(* IEC 61131-3 sources: BODAS-HelloWorld/st/bodas_rc18_12_40/plc_logic/application/02_easyconfig/dsm_easyconfig/structure (part 2) *)

(* ---- dfc_bds_tiinrow0x8b02-DFC_bds_TiInRow0x8B02.st ---- *)
(* --- Interface --- *)
{attribute 'external_name' := 'cmp_rts_DFC_bds_TiInRow0x8B02'}
TYPE DFC_bds_TiInRow0x8B02 : STRUCT
		DTC            : UDINT := 16#8B0200;
		DFCid          : UINT  := 102;
		debounceMethod : USINT := TIME_IN_ROW;
	END_STRUCT
END_TYPE

(* ---- dfc_bds_tiinrow0x8b03-DFC_bds_TiInRow0x8B03.st ---- *)
(* --- Interface --- *)
{attribute 'external_name' := 'cmp_rts_DFC_bds_TiInRow0x8B03'}
TYPE DFC_bds_TiInRow0x8B03 : STRUCT
		DTC            : UDINT := 16#8B0300;
		DFCid          : UINT  := 103;
		debounceMethod : USINT := TIME_IN_ROW;
	END_STRUCT
END_TYPE

(* ---- dfc_bds_tiupdwn0x8a01-DFC_bds_TiUpDwn0x8A01.st ---- *)
(* --- Interface --- *)
{attribute 'external_name' := 'cmp_rts_DFC_bds_TiUpDwn0x8A01'}
TYPE DFC_bds_TiUpDwn0x8A01 : STRUCT
		DTC            : UDINT := 16#8A0100;
		DFCid          : UINT  := 206;
		debounceMethod : USINT := TIME_UP_DOWN;
	END_STRUCT
END_TYPE

(* ---- dfc_bds_tiupdwn0x8a02-DFC_bds_TiUpDwn0x8A02.st ---- *)
(* --- Interface --- *)
{attribute 'external_name' := 'cmp_rts_DFC_bds_TiUpDwn0x8A02'}
TYPE DFC_bds_TiUpDwn0x8A02 : STRUCT
		DTC            : UDINT := 16#8A0200;
		DFCid          : UINT  := 207;
		debounceMethod : USINT := TIME_UP_DOWN;
	END_STRUCT
END_TYPE

(* ---- dfc_bds_tiupdwn0x8a03-DFC_bds_TiUpDwn0x8A03.st ---- *)
(* --- Interface --- *)
{attribute 'external_name' := 'cmp_rts_DFC_bds_TiUpDwn0x8A03'}
TYPE DFC_bds_TiUpDwn0x8A03 : STRUCT
		DTC            : UDINT := 16#8A0300;
		DFCid          : UINT  := 208;
		debounceMethod : USINT := TIME_UP_DOWN;
	END_STRUCT
END_TYPE

(* ---- dfc_can_e_timeout-DFC_CAN_E_TIMEOUT.st ---- *)
(* --- Interface --- *)
{attribute 'external_name' := 'cmp_rts_DFC_CAN_E_TIMEOUT'}
TYPE DFC_CAN_E_TIMEOUT : STRUCT
		DTC            : UDINT := 16#094200;
		DFCid          : UINT  := 1165;
		debounceMethod : USINT := NO_DEBOUNCE;
	END_STRUCT
END_TYPE

(* ---- dfc_cansm_e_bus_off_network_0-DFC_CANSM_E_BUS_OFF_NETWORK_0.st ---- *)
(* --- Interface --- *)
{attribute 'external_name' := 'cmp_rts_DFC_CANSM_E_BUS_OFF_NETWORK_0'}
TYPE DFC_CANSM_E_BUS_OFF_NETWORK_0 : STRUCT
		DTC            : UDINT := 16#104C00;
		DFCid          : UINT  := 1160;
		debounceMethod : USINT := NO_DEBOUNCE;
	END_STRUCT
END_TYPE

(* ---- dfc_cansm_e_bus_off_network_1-DFC_CANSM_E_BUS_OFF_NETWORK_1.st ---- *)
(* --- Interface --- *)
{attribute 'external_name' := 'cmp_rts_DFC_CANSM_E_BUS_OFF_NETWORK_1'}
TYPE DFC_CANSM_E_BUS_OFF_NETWORK_1 : STRUCT
		DTC            : UDINT := 16#104D00;
		DFCid          : UINT  := 1161;
		debounceMethod : USINT := NO_DEBOUNCE;
	END_STRUCT
END_TYPE

(* ---- dfc_cansm_e_bus_off_network_2-DFC_CANSM_E_BUS_OFF_NETWORK_2.st ---- *)
(* --- Interface --- *)
{attribute 'external_name' := 'cmp_rts_DFC_CANSM_E_BUS_OFF_NETWORK_2'}
TYPE DFC_CANSM_E_BUS_OFF_NETWORK_2 : STRUCT
		DTC            : UDINT := 16#104E00;
		DFCid          : UINT  := 1162;
		debounceMethod : USINT := NO_DEBOUNCE;
	END_STRUCT
END_TYPE

(* ---- dfc_cansm_e_bus_off_network_3-DFC_CANSM_E_BUS_OFF_NETWORK_3.st ---- *)
(* --- Interface --- *)
{attribute 'external_name' := 'cmp_rts_DFC_CANSM_E_BUS_OFF_NETWORK_3'}
TYPE DFC_CANSM_E_BUS_OFF_NETWORK_3 : STRUCT
		DTC            : UDINT := 16#104F00;
		DFCid          : UINT  := 1163;
		debounceMethod : USINT := NO_DEBOUNCE;
	END_STRUCT
END_TYPE

(* ---- dfc_cantrcv_e_no_trcv_control_0-DFC_CANTRCV_E_NO_TRCV_CONTROL_0.st ---- *)
(* --- Interface --- *)
{attribute 'external_name' := 'cmp_rts_DFC_CANTRCV_E_NO_TRCV_CONTROL_0'}
TYPE DFC_CANTRCV_E_NO_TRCV_CONTROL_0 : STRUCT
		DTC            : UDINT := 16#094000;
		DFCid          : UINT  := 1164;
		debounceMethod : USINT := NO_DEBOUNCE;
	END_STRUCT
END_TYPE

(* ---- dfc_com_numwhlincfrtleft-DFC_Com_numWhlIncFrtLeft.st ---- *)
(* --- Interface --- *)
{attribute 'external_name' := 'cmp_rts_DFC_Com_numWhlIncFrtLeft'}
TYPE DFC_Com_numWhlIncFrtLeft : STRUCT
		DTC : UDINT := 16#103A00;
	END_STRUCT
END_TYPE

(* ---- dfc_com_stwhlsensrrrht-DFC_Com_stWhlSensRrRht.st ---- *)
(* --- Interface --- *)
{attribute 'external_name' := 'cmp_rts_DFC_Com_stWhlSensRrRht'}
TYPE DFC_Com_stWhlSensRrRht : STRUCT
		DTC : UDINT := 16#103B00;
	END_STRUCT
END_TYPE

(* ---- dfc_com_trqclthtcsdcsdes-DFC_Com_trqClthTCSDCSDes.st ---- *)
(* --- Interface --- *)
{attribute 'external_name' := 'cmp_rts_DFC_Com_trqClthTCSDCSDes'}
TYPE DFC_Com_trqClthTCSDCSDes : STRUCT
		DTC : UDINT := 16#103C00;
	END_STRUCT
END_TYPE

(* ---- dfc_com_vwhlrrl-DFC_Com_vWhlRrL.st ---- *)
(* --- Interface --- *)
{attribute 'external_name' := 'cmp_rts_DFC_Com_vWhlRrL'}
TYPE DFC_Com_vWhlRrL : STRUCT
		DTC : UDINT := 16#103D00;
	END_STRUCT
END_TYPE

(* ---- dfc_comchksacc_06-DFC_ComChksACC_06.st ---- *)
(* --- Interface --- *)
{attribute 'external_name' := 'cmp_rts_DFC_ComChksACC_06'}
TYPE DFC_ComChksACC_06 : STRUCT
		DTC : UDINT := 16#101600;
	END_STRUCT
END_TYPE

(* ---- dfc_comchksbms_01-DFC_ComChksBMS_01.st ---- *)
(* --- Interface --- *)
{attribute 'external_name' := 'cmp_rts_DFC_ComChksBMS_01'}
TYPE DFC_ComChksBMS_01 : STRUCT
		DTC : UDINT := 16#101700;
	END_STRUCT
END_TYPE

(* ---- dfc_comchksesp_02-DFC_ComChksESP_02.st ---- *)
(* --- Interface --- *)
{attribute 'external_name' := 'cmp_rts_DFC_ComChksESP_02'}
TYPE DFC_ComChksESP_02 : STRUCT
		DTC : UDINT := 16#101800;
	END_STRUCT
END_TYPE

(* ---- dfc_comchksesp_05-DFC_ComChksESP_05.st ---- *)
(* --- Interface --- *)
{attribute 'external_name' := 'cmp_rts_DFC_ComChksESP_05'}
TYPE DFC_ComChksESP_05 : STRUCT
		DTC : UDINT := 16#101900;
	END_STRUCT
END_TYPE

(* ---- dfc_comchksesp_07-DFC_ComChksESP_07.st ---- *)
(* --- Interface --- *)
{attribute 'external_name' := 'cmp_rts_DFC_ComChksESP_07'}
TYPE DFC_ComChksESP_07 : STRUCT
		DTC : UDINT := 16#101A00;
	END_STRUCT
END_TYPE

(* ---- dfc_comchksesp_10-DFC_ComChksESP_10.st ---- *)
(* --- Interface --- *)
{attribute 'external_name' := 'cmp_rts_DFC_ComChksESP_10'}
TYPE DFC_ComChksESP_10 : STRUCT
		DTC : UDINT := 16#101B00;
	END_STRUCT
END_TYPE

(* ---- dfc_comchksesp_19-DFC_ComChksESP_19.st ---- *)
(* --- Interface --- *)
{attribute 'external_name' := 'cmp_rts_DFC_ComChksESP_19'}
TYPE DFC_ComChksESP_19 : STRUCT
		DTC : UDINT := 16#101C00;
	END_STRUCT
END_TYPE

(* ---- dfc_comchksesp_20-DFC_ComChksESP_20.st ---- *)
(* --- Interface --- *)
{attribute 'external_name' := 'cmp_rts_DFC_ComChksESP_20'}
TYPE DFC_ComChksESP_20 : STRUCT
		DTC : UDINT := 16#101D00;
	END_STRUCT
END_TYPE

(* ---- dfc_comchksesp_21-DFC_ComChksESP_21.st ---- *)
(* --- Interface --- *)
{attribute 'external_name' := 'cmp_rts_DFC_ComChksESP_21'}
TYPE DFC_ComChksESP_21 : STRUCT
		DTC : UDINT := 16#101E00;
	END_STRUCT
END_TYPE

(* ---- dfc_comchksklemmen_status_01-DFC_ComChksKlemmen_Status_01.st ---- *)
(* --- Interface --- *)
{attribute 'external_name' := 'cmp_rts_DFC_ComChksKlemmen_Status_01'}
TYPE DFC_ComChksKlemmen_Status_01 : STRUCT
		DTC : UDINT := 16#103800;
	END_STRUCT
END_TYPE

(* ---- dfc_comcntacc_06-DFC_ComCntACC_06.st ---- *)
(* --- Interface --- *)
{attribute 'external_name' := 'cmp_rts_DFC_ComCntACC_06'}
TYPE DFC_ComCntACC_06 : STRUCT
		DTC : UDINT := 16#101F00;
	END_STRUCT
END_TYPE

(* ---- dfc_comcntbms_01-DFC_ComCntBMS_01.st ---- *)
(* --- Interface --- *)
{attribute 'external_name' := 'cmp_rts_DFC_ComCntBMS_01'}
TYPE DFC_ComCntBMS_01 : STRUCT
		DTC : UDINT := 16#102000;
	END_STRUCT
END_TYPE

(* ---- dfc_comcntesp_02-DFC_ComCntESP_02.st ---- *)
(* --- Interface --- *)
{attribute 'external_name' := 'cmp_rts_DFC_ComCntESP_02'}
TYPE DFC_ComCntESP_02 : STRUCT
		DTC : UDINT := 16#102100;
	END_STRUCT
END_TYPE

(* ---- dfc_comcntesp_05-DFC_ComCntESP_05.st ---- *)
(* --- Interface --- *)
{attribute 'external_name' := 'cmp_rts_DFC_ComCntESP_05'}
TYPE DFC_ComCntESP_05 : STRUCT
		DTC : UDINT := 16#102200;
	END_STRUCT
END_TYPE

(* ---- dfc_comcntesp_07-DFC_ComCntESP_07.st ---- *)
(* --- Interface --- *)
{attribute 'external_name' := 'cmp_rts_DFC_ComCntESP_07'}
TYPE DFC_ComCntESP_07 : STRUCT
		DTC : UDINT := 16#102300;
	END_STRUCT
END_TYPE

(* ---- dfc_comcntesp_10-DFC_ComCntESP_10.st ---- *)
(* --- Interface --- *)
{attribute 'external_name' := 'cmp_rts_DFC_ComCntESP_10'}
TYPE DFC_ComCntESP_10 : STRUCT
		DTC : UDINT := 16#102400;
	END_STRUCT
END_TYPE

(* ---- dfc_comcntesp_19-DFC_ComCntESP_19.st ---- *)
(* --- Interface --- *)
{attribute 'external_name' := 'cmp_rts_DFC_ComCntESP_19'}
TYPE DFC_ComCntESP_19 : STRUCT
		DTC : UDINT := 16#102500;
	END_STRUCT
END_TYPE

(* ---- dfc_comcntesp_20-DFC_ComCntESP_20.st ---- *)
(* --- Interface --- *)
{attribute 'external_name' := 'cmp_rts_DFC_ComCntESP_20'}
TYPE DFC_ComCntESP_20 : STRUCT
		DTC : UDINT := 16#102600;
	END_STRUCT
END_TYPE

(* ---- dfc_comcntesp_21-DFC_ComCntESP_21.st ---- *)
(* --- Interface --- *)
{attribute 'external_name' := 'cmp_rts_DFC_ComCntESP_21'}
TYPE DFC_ComCntESP_21 : STRUCT
		DTC : UDINT := 16#102700;
	END_STRUCT
END_TYPE

(* ---- dfc_comcntklemmen_status_01-DFC_ComCntKlemmen_Status_01.st ---- *)
(* --- Interface --- *)
{attribute 'external_name' := 'cmp_rts_DFC_ComCntKlemmen_Status_01'}
TYPE DFC_ComCntKlemmen_Status_01 : STRUCT
		DTC : UDINT := 16#103900;
	END_STRUCT
END_TYPE

(* ---- dfc_comdlcacc_06-DFC_ComDlcACC_06.st ---- *)
(* --- Interface --- *)
{attribute 'external_name' := 'cmp_rts_DFC_ComDlcACC_06'}
TYPE DFC_ComDlcACC_06 : STRUCT
		DTC : UDINT := 16#102800;
	END_STRUCT
END_TYPE

(* ---- dfc_comdlcesp_02-DFC_ComDlcESP_02.st ---- *)
(* --- Interface --- *)
{attribute 'external_name' := 'cmp_rts_DFC_ComDlcESP_02'}
TYPE DFC_ComDlcESP_02 : STRUCT
		DTC : UDINT := 16#102900;
	END_STRUCT
END_TYPE

(* ---- dfc_comdlcesp_05-DFC_ComDlcESP_05.st ---- *)
(* --- Interface --- *)
{attribute 'external_name' := 'cmp_rts_DFC_ComDlcESP_05'}
TYPE DFC_ComDlcESP_05 : STRUCT
		DTC : UDINT := 16#102A00;
	END_STRUCT
END_TYPE

(* ---- dfc_comdlcesp_07-DFC_ComDlcESP_07.st ---- *)
(* --- Interface --- *)
{attribute 'external_name' := 'cmp_rts_DFC_ComDlcESP_07'}
TYPE DFC_ComDlcESP_07 : STRUCT
		DTC : UDINT := 16#102B00;
	END_STRUCT
END_TYPE

(* ---- dfc_comdlcesp_10-DFC_ComDlcESP_10.st ---- *)
(* --- Interface --- *)
{attribute 'external_name' := 'cmp_rts_DFC_ComDlcESP_10'}
TYPE DFC_ComDlcESP_10 : STRUCT
		DTC : UDINT := 16#102C00;
	END_STRUCT
END_TYPE

(* ---- dfc_comdlcesp_19-DFC_ComDlcESP_19.st ---- *)
(* --- Interface --- *)
{attribute 'external_name' := 'cmp_rts_DFC_ComDlcESP_19'}
TYPE DFC_ComDlcESP_19 : STRUCT
		DTC : UDINT := 16#102D00;
	END_STRUCT
END_TYPE

(* ---- dfc_comdlcesp_20-DFC_ComDlcESP_20.st ---- *)
(* --- Interface --- *)
{attribute 'external_name' := 'cmp_rts_DFC_ComDlcESP_20'}
TYPE DFC_ComDlcESP_20 : STRUCT
		DTC : UDINT := 16#102E00;
	END_STRUCT
END_TYPE

(* ---- dfc_comdlcesp_21-DFC_ComDlcESP_21.st ---- *)
(* --- Interface --- *)
{attribute 'external_name' := 'cmp_rts_DFC_ComDlcESP_21'}
TYPE DFC_ComDlcESP_21 : STRUCT
		DTC : UDINT := 16#102F00;
	END_STRUCT
END_TYPE

(* ---- dfc_comm_e_net_start_ind_channel_0-DFC_COMM_E_NET_START_IND_CHANNEL_0.st ---- *)
(* --- Interface --- *)
{attribute 'external_name' := 'cmp_rts_DFC_COMM_E_NET_START_IND_CHANNEL_0'}
TYPE DFC_COMM_E_NET_START_IND_CHANNEL_0 : STRUCT
		DTC            : UDINT := 16#105000;
		DFCid          : UINT  := 1166;
		debounceMethod : USINT := NO_DEBOUNCE;
	END_STRUCT
END_TYPE

(* ---- dfc_comm_e_net_start_ind_channel_1-DFC_COMM_E_NET_START_IND_CHANNEL_1.st ---- *)
(* --- Interface --- *)
{attribute 'external_name' := 'cmp_rts_DFC_COMM_E_NET_START_IND_CHANNEL_1'}
TYPE DFC_COMM_E_NET_START_IND_CHANNEL_1 : STRUCT
		DTC            : UDINT := 16#105100;
		DFCid          : UINT  := 1167;
		debounceMethod : USINT := NO_DEBOUNCE;
	END_STRUCT
END_TYPE

(* ---- dfc_comm_e_net_start_ind_channel_2-DFC_COMM_E_NET_START_IND_CHANNEL_2.st ---- *)
(* --- Interface --- *)
{attribute 'external_name' := 'cmp_rts_DFC_COMM_E_NET_START_IND_CHANNEL_2'}
TYPE DFC_COMM_E_NET_START_IND_CHANNEL_2 : STRUCT
		DTC            : UDINT := 16#105200;
		DFCid          : UINT  := 1168;
		debounceMethod : USINT := NO_DEBOUNCE;
	END_STRUCT
END_TYPE

(* ---- dfc_comm_e_net_start_ind_channel_3-DFC_COMM_E_NET_START_IND_CHANNEL_3.st ---- *)
(* --- Interface --- *)
{attribute 'external_name' := 'cmp_rts_DFC_COMM_E_NET_START_IND_CHANNEL_3'}
TYPE DFC_COMM_E_NET_START_IND_CHANNEL_3 : STRUCT
		DTC            : UDINT := 16#105300;
		DFCid          : UINT  := 1169;
		debounceMethod : USINT := NO_DEBOUNCE;
	END_STRUCT
END_TYPE

(* ---- dfc_comm_e_net_start_ind_channel_4-DFC_COMM_E_NET_START_IND_CHANNEL_4.st ---- *)
(* --- Interface --- *)
{attribute 'external_name' := 'cmp_rts_DFC_COMM_E_NET_START_IND_CHANNEL_4'}
TYPE DFC_COMM_E_NET_START_IND_CHANNEL_4 : STRUCT
		DTC            : UDINT := 16#105400;
		DFCid          : UINT  := 1170;
		debounceMethod : USINT := NO_DEBOUNCE;
	END_STRUCT
END_TYPE

(* ---- dfc_comm_e_net_start_ind_channel_5-DFC_COMM_E_NET_START_IND_CHANNEL_5.st ---- *)
(* --- Interface --- *)
{attribute 'external_name' := 'cmp_rts_DFC_COMM_E_NET_START_IND_CHANNEL_5'}
TYPE DFC_COMM_E_NET_START_IND_CHANNEL_5 : STRUCT
		DTC            : UDINT := 16#105500;
		DFCid          : UINT  := 1171;
		debounceMethod : USINT := NO_DEBOUNCE;
	END_STRUCT
END_TYPE

(* ---- dfc_comtoutacc_06-DFC_ComTOutACC_06.st ---- *)
(* --- Interface --- *)
{attribute 'external_name' := 'cmp_rts_DFC_ComTOutACC_06'}
TYPE DFC_ComTOutACC_06 : STRUCT
		DTC : UDINT := 16#103000;
	END_STRUCT
END_TYPE

(* ---- dfc_comtoutesp_02-DFC_ComTOutESP_02.st ---- *)
(* --- Interface --- *)
{attribute 'external_name' := 'cmp_rts_DFC_ComTOutESP_02'}
TYPE DFC_ComTOutESP_02 : STRUCT
		DTC : UDINT := 16#103100;
	END_STRUCT
END_TYPE

(* ---- dfc_comtoutesp_05-DFC_ComTOutESP_05.st ---- *)
(* --- Interface --- *)
{attribute 'external_name' := 'cmp_rts_DFC_ComTOutESP_05'}
TYPE DFC_ComTOutESP_05 : STRUCT
		DTC : UDINT := 16#103200;
	END_STRUCT
END_TYPE

(* ---- dfc_comtoutesp_07-DFC_ComTOutESP_07.st ---- *)
(* --- Interface --- *)
{attribute 'external_name' := 'cmp_rts_DFC_ComTOutESP_07'}
TYPE DFC_ComTOutESP_07 : STRUCT
		DTC : UDINT := 16#103300;
	END_STRUCT
END_TYPE

(* ---- dfc_comtoutesp_10-DFC_ComTOutESP_10.st ---- *)
(* --- Interface --- *)
{attribute 'external_name' := 'cmp_rts_DFC_ComTOutESP_10'}
TYPE DFC_ComTOutESP_10 : STRUCT
		DTC : UDINT := 16#103400;
	END_STRUCT
END_TYPE

(* ---- dfc_comtoutesp_19-DFC_ComTOutESP_19.st ---- *)
(* --- Interface --- *)
{attribute 'external_name' := 'cmp_rts_DFC_ComTOutESP_19'}
TYPE DFC_ComTOutESP_19 : STRUCT
		DTC : UDINT := 16#103500;
	END_STRUCT
END_TYPE

(* ---- dfc_comtoutesp_20-DFC_ComTOutESP_20.st ---- *)
(* --- Interface --- *)
{attribute 'external_name' := 'cmp_rts_DFC_ComTOutESP_20'}
TYPE DFC_ComTOutESP_20 : STRUCT
		DTC : UDINT := 16#103600;
	END_STRUCT
END_TYPE

(* ---- dfc_comtoutesp_21-DFC_ComTOutESP_21.st ---- *)
(* --- Interface --- *)
{attribute 'external_name' := 'cmp_rts_DFC_ComTOutESP_21'}
TYPE DFC_ComTOutESP_21 : STRUCT
		DTC : UDINT := 16#103700;
	END_STRUCT
END_TYPE

(* ---- dfc_devlibbattuhi-DFC_DevLibBattUHi.st ---- *)
(* --- Interface --- *)
{attribute 'external_name' := 'cmp_rts_DFC_DevLibBattUHi'}
TYPE DFC_DevLibBattUHi : STRUCT
		DTC            : UDINT := 16#092300;
		DFCid          : UINT  := 104;
		debounceMethod : USINT := TIME_UP_DOWN;
	END_STRUCT
END_TYPE

(* ---- dfc_devlibbattulo-DFC_DevLibBattULo.st ---- *)
(* --- Interface --- *)
{attribute 'external_name' := 'cmp_rts_DFC_DevLibBattULo'}
TYPE DFC_DevLibBattULo : STRUCT
		DTC            : UDINT := 16#092400;
		DFCid          : UINT  := 105;
		debounceMethod : USINT := TIME_UP_DOWN;
	END_STRUCT
END_TYPE

(* ---- dfc_dsmdummy-DFC_DSMDummy.st ---- *)
(* --- Interface --- *)
{attribute 'external_name' := 'cmp_rts_DFC_DSMDummy'}
TYPE DFC_DSMDummy : STRUCT
		DTC            : UDINT := 16#100F00;
		DFCid          : UINT  := 720;
		debounceMethod : USINT := NO_DEBOUNCE;
	END_STRUCT
END_TYPE

(* ---- dfc_lin_e_timeout-DFC_LIN_E_TIMEOUT.st ---- *)
(* --- Interface --- *)
{attribute 'external_name' := 'cmp_rts_DFC_LIN_E_TIMEOUT'}
TYPE DFC_LIN_E_TIMEOUT : STRUCT
		DTC            : UDINT := 16#094100;
		DFCid          : UINT  := 1172;
		debounceMethod : USINT := NO_DEBOUNCE;
	END_STRUCT
END_TYPE

(* ---- dfc_mocsopico-DFC_MoCSOPICO.st ---- *)
(* --- Interface --- *)
{attribute 'external_name' := 'cmp_rts_DFC_MoCSOPICO'}
TYPE DFC_MoCSOPICO : STRUCT
		DTC            : UDINT := 16#106000;
		DFCid          : UINT  := 1296;
		debounceMethod : USINT := NATIVE;
	END_STRUCT
END_TYPE

(* ---- dfc_mofvarpostbldsel-DFC_MoFVarPostBldSel.st ---- *)
(* --- Interface --- *)
{attribute 'external_name' := 'cmp_rts_DFC_MoFVarPostBldSel'}
TYPE DFC_MoFVarPostBldSel : STRUCT
		DTC            : UDINT := 16#098900;
		DFCid          : UINT  := 1297;
		debounceMethod : USINT := NATIVE;
	END_STRUCT
END_TYPE

(* ---- dfc_mosysctrlreini-DFC_MoSysCtrlReIni.st ---- *)
(* --- Interface --- *)
{attribute 'external_name' := 'cmp_rts_DFC_MoSysCtrlReIni'}
TYPE DFC_MoSysCtrlReIni : STRUCT
		DTC            : UDINT := 16#106100;
		DFCid          : UINT  := 1298;
		debounceMethod : USINT := NATIVE;
	END_STRUCT
END_TYPE

(* ---- dfc_moxemm_smu_alm0_0-DFC_MOXEMM_SMU_ALM0_0.st ---- *)
(* --- Interface --- *)
{attribute 'external_name' := 'cmp_rts_DFC_MOXEMM_SMU_ALM0_0'}
TYPE DFC_MOXEMM_SMU_ALM0_0 : STRUCT
		DTC            : UDINT := 16#106200;
		DFCid          : UINT  := 1185;
		debounceMethod : USINT := NATIVE;
	END_STRUCT
END_TYPE

(* ---- dfc_moxemm_smu_alm0_1-DFC_MOXEMM_SMU_ALM0_1.st ---- *)
(* --- Interface --- *)
{attribute 'external_name' := 'cmp_rts_DFC_MOXEMM_SMU_ALM0_1'}
TYPE DFC_MOXEMM_SMU_ALM0_1 : STRUCT
		DTC            : UDINT := 16#106300;
		DFCid          : UINT  := 1186;
		debounceMethod : USINT := NATIVE;
	END_STRUCT
END_TYPE

(* ---- dfc_moxemm_smu_alm0_10-DFC_MOXEMM_SMU_ALM0_10.st ---- *)
(* --- Interface --- *)
{attribute 'external_name' := 'cmp_rts_DFC_MOXEMM_SMU_ALM0_10'}
TYPE DFC_MOXEMM_SMU_ALM0_10 : STRUCT
		DTC            : UDINT := 16#106900;
		DFCid          : UINT  := 1187;
		debounceMethod : USINT := NATIVE;
	END_STRUCT
END_TYPE

(* ---- dfc_moxemm_smu_alm0_11-DFC_MOXEMM_SMU_ALM0_11.st ---- *)
(* --- Interface --- *)
{attribute 'external_name' := 'cmp_rts_DFC_MOXEMM_SMU_ALM0_11'}
TYPE DFC_MOXEMM_SMU_ALM0_11 : STRUCT
		DTC            : UDINT := 16#106A00;
		DFCid          : UINT  := 1188;
		debounceMethod : USINT := NATIVE;
	END_STRUCT
END_TYPE

(* ---- dfc_moxemm_smu_alm0_13-DFC_MOXEMM_SMU_ALM0_13.st ---- *)
(* --- Interface --- *)
{attribute 'external_name' := 'cmp_rts_DFC_MOXEMM_SMU_ALM0_13'}
TYPE DFC_MOXEMM_SMU_ALM0_13 : STRUCT
		DTC            : UDINT := 16#106B00;
		DFCid          : UINT  := 1189;
		debounceMethod : USINT := NATIVE;
	END_STRUCT
END_TYPE

(* ---- dfc_moxemm_smu_alm0_14-DFC_MOXEMM_SMU_ALM0_14.st ---- *)
(* --- Interface --- *)
{attribute 'external_name' := 'cmp_rts_DFC_MOXEMM_SMU_ALM0_14'}
TYPE DFC_MOXEMM_SMU_ALM0_14 : STRUCT
		DTC            : UDINT := 16#106C00;
		DFCid          : UINT  := 1190;
		debounceMethod : USINT := NATIVE;
	END_STRUCT
END_TYPE

(* ---- dfc_moxemm_smu_alm0_2-DFC_MOXEMM_SMU_ALM0_2.st ---- *)
(* --- Interface --- *)
{attribute 'external_name' := 'cmp_rts_DFC_MOXEMM_SMU_ALM0_2'}
TYPE DFC_MOXEMM_SMU_ALM0_2 : STRUCT
		DTC            : UDINT := 16#106400;
		DFCid          : UINT  := 1191;
		debounceMethod : USINT := NATIVE;
	END_STRUCT
END_TYPE

(* ---- dfc_moxemm_smu_alm0_22-DFC_MOXEMM_SMU_ALM0_22.st ---- *)
(* --- Interface --- *)
{attribute 'external_name' := 'cmp_rts_DFC_MOXEMM_SMU_ALM0_22'}
TYPE DFC_MOXEMM_SMU_ALM0_22 : STRUCT
		DTC            : UDINT := 16#106D00;
		DFCid          : UINT  := 1192;
		debounceMethod : USINT := NATIVE;
	END_STRUCT
END_TYPE

(* ---- dfc_moxemm_smu_alm0_23-DFC_MOXEMM_SMU_ALM0_23.st ---- *)
(* --- Interface --- *)
{attribute 'external_name' := 'cmp_rts_DFC_MOXEMM_SMU_ALM0_23'}
TYPE DFC_MOXEMM_SMU_ALM0_23 : STRUCT
		DTC            : UDINT := 16#106E00;
		DFCid          : UINT  := 1193;
		debounceMethod : USINT := NATIVE;
	END_STRUCT
END_TYPE

(* ---- dfc_moxemm_smu_alm0_4-DFC_MOXEMM_SMU_ALM0_4.st ---- *)
(* --- Interface --- *)
{attribute 'external_name' := 'cmp_rts_DFC_MOXEMM_SMU_ALM0_4'}
TYPE DFC_MOXEMM_SMU_ALM0_4 : STRUCT
		DTC            : UDINT := 16#106500;
		DFCid          : UINT  := 1194;
		debounceMethod : USINT := NATIVE;
	END_STRUCT
END_TYPE

(* ---- dfc_moxemm_smu_alm0_5-DFC_MOXEMM_SMU_ALM0_5.st ---- *)
(* --- Interface --- *)
{attribute 'external_name' := 'cmp_rts_DFC_MOXEMM_SMU_ALM0_5'}
TYPE DFC_MOXEMM_SMU_ALM0_5 : STRUCT
		DTC            : UDINT := 16#106600;
		DFCid          : UINT  := 1195;
		debounceMethod : USINT := NATIVE;
	END_STRUCT
END_TYPE

(* ---- dfc_moxemm_smu_alm0_7-DFC_MOXEMM_SMU_ALM0_7.st ---- *)
(* --- Interface --- *)
{attribute 'external_name' := 'cmp_rts_DFC_MOXEMM_SMU_ALM0_7'}
TYPE DFC_MOXEMM_SMU_ALM0_7 : STRUCT
		DTC            : UDINT := 16#106700;
		DFCid          : UINT  := 1196;
		debounceMethod : USINT := NATIVE;
	END_STRUCT
END_TYPE

(* ---- dfc_moxemm_smu_alm0_8-DFC_MOXEMM_SMU_ALM0_8.st ---- *)
(* --- Interface --- *)
{attribute 'external_name' := 'cmp_rts_DFC_MOXEMM_SMU_ALM0_8'}
TYPE DFC_MOXEMM_SMU_ALM0_8 : STRUCT
		DTC            : UDINT := 16#106800;
		DFCid          : UINT  := 1197;
		debounceMethod : USINT := NATIVE;
	END_STRUCT
END_TYPE

(* ---- dfc_moxemm_smu_alm10_16-DFC_MOXEMM_SMU_ALM10_16.st ---- *)
(* --- Interface --- *)
{attribute 'external_name' := 'cmp_rts_DFC_MOXEMM_SMU_ALM10_16'}
TYPE DFC_MOXEMM_SMU_ALM10_16 : STRUCT
		DTC            : UDINT := 16#10C200;
		DFCid          : UINT  := 1198;
		debounceMethod : USINT := NATIVE;
	END_STRUCT
END_TYPE

(* ---- dfc_moxemm_smu_alm10_17-DFC_MOXEMM_SMU_ALM10_17.st ---- *)
(* --- Interface --- *)
{attribute 'external_name' := 'cmp_rts_DFC_MOXEMM_SMU_ALM10_17'}
TYPE DFC_MOXEMM_SMU_ALM10_17 : STRUCT
		DTC            : UDINT := 16#10C300;
		DFCid          : UINT  := 1199;
		debounceMethod : USINT := NATIVE;
	END_STRUCT
END_TYPE

(* ---- dfc_moxemm_smu_alm10_21-DFC_MOXEMM_SMU_ALM10_21.st ---- *)
(* --- Interface --- *)
{attribute 'external_name' := 'cmp_rts_DFC_MOXEMM_SMU_ALM10_21'}
TYPE DFC_MOXEMM_SMU_ALM10_21 : STRUCT
		DTC            : UDINT := 16#10C400;
		DFCid          : UINT  := 1200;
		debounceMethod : USINT := NATIVE;
	END_STRUCT
END_TYPE

(* ---- dfc_moxemm_smu_alm11_0-DFC_MOXEMM_SMU_ALM11_0.st ---- *)
(* --- Interface --- *)
{attribute 'external_name' := 'cmp_rts_DFC_MOXEMM_SMU_ALM11_0'}
TYPE DFC_MOXEMM_SMU_ALM11_0 : STRUCT
		DTC            : UDINT := 16#10C500;
		DFCid          : UINT  := 1201;
		debounceMethod : USINT := NATIVE;
	END_STRUCT
END_TYPE

(* ---- dfc_moxemm_smu_alm11_1-DFC_MOXEMM_SMU_ALM11_1.st ---- *)
(* --- Interface --- *)
{attribute 'external_name' := 'cmp_rts_DFC_MOXEMM_SMU_ALM11_1'}
TYPE DFC_MOXEMM_SMU_ALM11_1 : STRUCT
		DTC            : UDINT := 16#10C600;
		DFCid          : UINT  := 1202;
		debounceMethod : USINT := NATIVE;
	END_STRUCT
END_TYPE

(* ---- dfc_moxemm_smu_alm11_2-DFC_MOXEMM_SMU_ALM11_2.st ---- *)
(* --- Interface --- *)
{attribute 'external_name' := 'cmp_rts_DFC_MOXEMM_SMU_ALM11_2'}
TYPE DFC_MOXEMM_SMU_ALM11_2 : STRUCT
		DTC            : UDINT := 16#10C700;
		DFCid          : UINT  := 1203;
		debounceMethod : USINT := NATIVE;
	END_STRUCT
END_TYPE

(* ---- dfc_moxemm_smu_alm11_3-DFC_MOXEMM_SMU_ALM11_3.st ---- *)
(* --- Interface --- *)
{attribute 'external_name' := 'cmp_rts_DFC_MOXEMM_SMU_ALM11_3'}
TYPE DFC_MOXEMM_SMU_ALM11_3 : STRUCT
		DTC            : UDINT := 16#10C800;
		DFCid          : UINT  := 1204;
		debounceMethod : USINT := NATIVE;
	END_STRUCT
END_TYPE

(* ---- dfc_moxemm_smu_alm11_4-DFC_MOXEMM_SMU_ALM11_4.st ---- *)
(* --- Interface --- *)
{attribute 'external_name' := 'cmp_rts_DFC_MOXEMM_SMU_ALM11_4'}
TYPE DFC_MOXEMM_SMU_ALM11_4 : STRUCT
		DTC            : UDINT := 16#10C900;
		DFCid          : UINT  := 1205;
		debounceMethod : USINT := NATIVE;
	END_STRUCT
END_TYPE

(* ---- dfc_moxemm_smu_alm11_5-DFC_MOXEMM_SMU_ALM11_5.st ---- *)
(* --- Interface --- *)
{attribute 'external_name' := 'cmp_rts_DFC_MOXEMM_SMU_ALM11_5'}
TYPE DFC_MOXEMM_SMU_ALM11_5 : STRUCT
		DTC            : UDINT := 16#10CA00;
		DFCid          : UINT  := 1206;
		debounceMethod : USINT := NATIVE;
	END_STRUCT
END_TYPE

(* ---- dfc_moxemm_smu_alm11_8-DFC_MOXEMM_SMU_ALM11_8.st ---- *)
(* --- Interface --- *)
{attribute 'external_name' := 'cmp_rts_DFC_MOXEMM_SMU_ALM11_8'}
TYPE DFC_MOXEMM_SMU_ALM11_8 : STRUCT
		DTC            : UDINT := 16#10CB00;
		DFCid          : UINT  := 1207;
		debounceMethod : USINT := NATIVE;
	END_STRUCT
END_TYPE

(* ---- dfc_moxemm_smu_alm11_9-DFC_MOXEMM_SMU_ALM11_9.st ---- *)
(* --- Interface --- *)
{attribute 'external_name' := 'cmp_rts_DFC_MOXEMM_SMU_ALM11_9'}
TYPE DFC_MOXEMM_SMU_ALM11_9 : STRUCT
		DTC            : UDINT := 16#10CC00;
		DFCid          : UINT  := 1208;
		debounceMethod : USINT := NATIVE;
	END_STRUCT
END_TYPE

(* ---- dfc_moxemm_smu_alm1_0-DFC_MOXEMM_SMU_ALM1_0.st ---- *)
(* --- Interface --- *)
{attribute 'external_name' := 'cmp_rts_DFC_MOXEMM_SMU_ALM1_0'}
TYPE DFC_MOXEMM_SMU_ALM1_0 : STRUCT
		DTC            : UDINT := 16#106F00;
		DFCid          : UINT  := 1209;
		debounceMethod : USINT := NATIVE;
	END_STRUCT
END_TYPE

(* ---- dfc_moxemm_smu_alm1_1-DFC_MOXEMM_SMU_ALM1_1.st ---- *)
(* --- Interface --- *)
{attribute 'external_name' := 'cmp_rts_DFC_MOXEMM_SMU_ALM1_1'}
TYPE DFC_MOXEMM_SMU_ALM1_1 : STRUCT
		DTC            : UDINT := 16#107000;
		DFCid          : UINT  := 1210;
		debounceMethod : USINT := NATIVE;
	END_STRUCT
END_TYPE

(* ---- dfc_moxemm_smu_alm1_10-DFC_MOXEMM_SMU_ALM1_10.st ---- *)
(* --- Interface --- *)
{attribute 'external_name' := 'cmp_rts_DFC_MOXEMM_SMU_ALM1_10'}
TYPE DFC_MOXEMM_SMU_ALM1_10 : STRUCT
		DTC            : UDINT := 16#107600;
		DFCid          : UINT  := 1211;
		debounceMethod : USINT := NATIVE;
	END_STRUCT
END_TYPE

(* ---- dfc_moxemm_smu_alm1_11-DFC_MOXEMM_SMU_ALM1_11.st ---- *)
(* --- Interface --- *)
{attribute 'external_name' := 'cmp_rts_DFC_MOXEMM_SMU_ALM1_11'}
TYPE DFC_MOXEMM_SMU_ALM1_11 : STRUCT
		DTC            : UDINT := 16#107700;
		DFCid          : UINT  := 1212;
		debounceMethod : USINT := NATIVE;
	END_STRUCT
END_TYPE

(* ---- dfc_moxemm_smu_alm1_13-DFC_MOXEMM_SMU_ALM1_13.st ---- *)
(* --- Interface --- *)
{attribute 'external_name' := 'cmp_rts_DFC_MOXEMM_SMU_ALM1_13'}
TYPE DFC_MOXEMM_SMU_ALM1_13 : STRUCT
		DTC            : UDINT := 16#107800;
		DFCid          : UINT  := 1213;
		debounceMethod : USINT := NATIVE;
	END_STRUCT
END_TYPE

(* ---- dfc_moxemm_smu_alm1_14-DFC_MOXEMM_SMU_ALM1_14.st ---- *)
(* --- Interface --- *)
{attribute 'external_name' := 'cmp_rts_DFC_MOXEMM_SMU_ALM1_14'}
TYPE DFC_MOXEMM_SMU_ALM1_14 : STRUCT
		DTC            : UDINT := 16#107900;
		DFCid          : UINT  := 1214;
		debounceMethod : USINT := NATIVE;
	END_STRUCT
END_TYPE

(* ---- dfc_moxemm_smu_alm1_2-DFC_MOXEMM_SMU_ALM1_2.st ---- *)
(* --- Interface --- *)
{attribute 'external_name' := 'cmp_rts_DFC_MOXEMM_SMU_ALM1_2'}
TYPE DFC_MOXEMM_SMU_ALM1_2 : STRUCT
		DTC            : UDINT := 16#107100;
		DFCid          : UINT  := 1215;
		debounceMethod : USINT := NATIVE;
	END_STRUCT
END_TYPE

(* ---- dfc_moxemm_smu_alm1_22-DFC_MOXEMM_SMU_ALM1_22.st ---- *)
(* --- Interface --- *)
{attribute 'external_name' := 'cmp_rts_DFC_MOXEMM_SMU_ALM1_22'}
TYPE DFC_MOXEMM_SMU_ALM1_22 : STRUCT
		DTC            : UDINT := 16#107A00;
		DFCid          : UINT  := 1216;
		debounceMethod : USINT := NATIVE;
	END_STRUCT
END_TYPE

(* ---- dfc_moxemm_smu_alm1_23-DFC_MOXEMM_SMU_ALM1_23.st ---- *)
(* --- Interface --- *)
{attribute 'external_name' := 'cmp_rts_DFC_MOXEMM_SMU_ALM1_23'}
TYPE DFC_MOXEMM_SMU_ALM1_23 : STRUCT
		DTC            : UDINT := 16#107B00;
		DFCid          : UINT  := 1217;
		debounceMethod : USINT := NATIVE;
	END_STRUCT
END_TYPE

(* ---- dfc_moxemm_smu_alm1_4-DFC_MOXEMM_SMU_ALM1_4.st ---- *)
(* --- Interface --- *)
{attribute 'external_name' := 'cmp_rts_DFC_MOXEMM_SMU_ALM1_4'}
TYPE DFC_MOXEMM_SMU_ALM1_4 : STRUCT
		DTC            : UDINT := 16#107200;
		DFCid          : UINT  := 1218;
		debounceMethod : USINT := NATIVE;
	END_STRUCT
END_TYPE

(* ---- dfc_moxemm_smu_alm1_5-DFC_MOXEMM_SMU_ALM1_5.st ---- *)
(* --- Interface --- *)
{attribute 'external_name' := 'cmp_rts_DFC_MOXEMM_SMU_ALM1_5'}
TYPE DFC_MOXEMM_SMU_ALM1_5 : STRUCT
		DTC            : UDINT := 16#107300;
		DFCid          : UINT  := 1219;
		debounceMethod : USINT := NATIVE;
	END_STRUCT
END_TYPE

(* ---- dfc_moxemm_smu_alm1_7-DFC_MOXEMM_SMU_ALM1_7.st ---- *)
(* --- Interface --- *)
{attribute 'external_name' := 'cmp_rts_DFC_MOXEMM_SMU_ALM1_7'}
TYPE DFC_MOXEMM_SMU_ALM1_7 : STRUCT
		DTC            : UDINT := 16#107400;
		DFCid          : UINT  := 1220;
		debounceMethod : USINT := NATIVE;
	END_STRUCT
END_TYPE

(* ---- dfc_moxemm_smu_alm1_8-DFC_MOXEMM_SMU_ALM1_8.st ---- *)
(* --- Interface --- *)
{attribute 'external_name' := 'cmp_rts_DFC_MOXEMM_SMU_ALM1_8'}
TYPE DFC_MOXEMM_SMU_ALM1_8 : STRUCT
		DTC            : UDINT := 16#107500;
		DFCid          : UINT  := 1221;
		debounceMethod : USINT := NATIVE;
	END_STRUCT
END_TYPE

(* ---- dfc_moxemm_smu_alm21_0-DFC_MOXEMM_SMU_ALM21_0.st ---- *)
(* --- Interface --- *)
{attribute 'external_name' := 'cmp_rts_DFC_MOXEMM_SMU_ALM21_0'}
TYPE DFC_MOXEMM_SMU_ALM21_0 : STRUCT
		DTC            : UDINT := 16#10CD00;
		DFCid          : UINT  := 1222;
		debounceMethod : USINT := NATIVE;
	END_STRUCT
END_TYPE

(* ---- dfc_moxemm_smu_alm21_16-DFC_MOXEMM_SMU_ALM21_16.st ---- *)
(* --- Interface --- *)
{attribute 'external_name' := 'cmp_rts_DFC_MOXEMM_SMU_ALM21_16'}
TYPE DFC_MOXEMM_SMU_ALM21_16 : STRUCT
		DTC            : UDINT := 16#10CF00;
		DFCid          : UINT  := 1223;
		debounceMethod : USINT := NATIVE;
	END_STRUCT
END_TYPE

(* ---- dfc_moxemm_smu_alm21_3-DFC_MOXEMM_SMU_ALM21_3.st ---- *)
(* --- Interface --- *)
{attribute 'external_name' := 'cmp_rts_DFC_MOXEMM_SMU_ALM21_3'}
TYPE DFC_MOXEMM_SMU_ALM21_3 : STRUCT
		DTC            : UDINT := 16#10CE00;
		DFCid          : UINT  := 1224;
		debounceMethod : USINT := NATIVE;
	END_STRUCT
END_TYPE

(* ---- dfc_moxemm_smu_alm2_1-DFC_MOXEMM_SMU_ALM2_1.st ---- *)
(* --- Interface --- *)
{attribute 'external_name' := 'cmp_rts_DFC_MOXEMM_SMU_ALM2_1'}
TYPE DFC_MOXEMM_SMU_ALM2_1 : STRUCT
		DTC            : UDINT := 16#107C00;
		DFCid          : UINT  := 1225;
		debounceMethod : USINT := NATIVE;
	END_STRUCT
END_TYPE

(* ---- dfc_moxemm_smu_alm2_10-DFC_MOXEMM_SMU_ALM2_10.st ---- *)
(* --- Interface --- *)
{attribute 'external_name' := 'cmp_rts_DFC_MOXEMM_SMU_ALM2_10'}
TYPE DFC_MOXEMM_SMU_ALM2_10 : STRUCT
		DTC            : UDINT := 16#108200;
		DFCid          : UINT  := 1226;
		debounceMethod : USINT := NATIVE;
	END_STRUCT
END_TYPE

(* ---- dfc_moxemm_smu_alm2_11-DFC_MOXEMM_SMU_ALM2_11.st ---- *)
(* --- Interface --- *)
{attribute 'external_name' := 'cmp_rts_DFC_MOXEMM_SMU_ALM2_11'}
TYPE DFC_MOXEMM_SMU_ALM2_11 : STRUCT
		DTC            : UDINT := 16#108300;
		DFCid          : UINT  := 1227;
		debounceMethod : USINT := NATIVE;
	END_STRUCT
END_TYPE

(* ---- dfc_moxemm_smu_alm2_13-DFC_MOXEMM_SMU_ALM2_13.st ---- *)
(* --- Interface --- *)
{attribute 'external_name' := 'cmp_rts_DFC_MOXEMM_SMU_ALM2_13'}
TYPE DFC_MOXEMM_SMU_ALM2_13 : STRUCT
		DTC            : UDINT := 16#108400;
		DFCid          : UINT  := 1228;
		debounceMethod : USINT := NATIVE;
	END_STRUCT
END_TYPE

(* ---- dfc_moxemm_smu_alm2_14-DFC_MOXEMM_SMU_ALM2_14.st ---- *)
(* --- Interface --- *)
{attribute 'external_name' := 'cmp_rts_DFC_MOXEMM_SMU_ALM2_14'}
TYPE DFC_MOXEMM_SMU_ALM2_14 : STRUCT
		DTC            : UDINT := 16#108500;
		DFCid          : UINT  := 1229;
		debounceMethod : USINT := NATIVE;
	END_STRUCT
END_TYPE

(* ---- dfc_moxemm_smu_alm2_2-DFC_MOXEMM_SMU_ALM2_2.st ---- *)
(* --- Interface --- *)
{attribute 'external_name' := 'cmp_rts_DFC_MOXEMM_SMU_ALM2_2'}
TYPE DFC_MOXEMM_SMU_ALM2_2 : STRUCT
		DTC            : UDINT := 16#107D00;
		DFCid          : UINT  := 1230;
		debounceMethod : USINT := NATIVE;
	END_STRUCT
END_TYPE

(* ---- dfc_moxemm_smu_alm2_22-DFC_MOXEMM_SMU_ALM2_22.st ---- *)
(* --- Interface --- *)
{attribute 'external_name' := 'cmp_rts_DFC_MOXEMM_SMU_ALM2_22'}
TYPE DFC_MOXEMM_SMU_ALM2_22 : STRUCT
		DTC            : UDINT := 16#108600;
		DFCid          : UINT  := 1231;
		debounceMethod : USINT := NATIVE;
	END_STRUCT
END_TYPE

(* ---- dfc_moxemm_smu_alm2_23-DFC_MOXEMM_SMU_ALM2_23.st ---- *)
(* --- Interface --- *)
{attribute 'external_name' := 'cmp_rts_DFC_MOXEMM_SMU_ALM2_23'}
TYPE DFC_MOXEMM_SMU_ALM2_23 : STRUCT
		DTC            : UDINT := 16#108700;
		DFCid          : UINT  := 1232;
		debounceMethod : USINT := NATIVE;
	END_STRUCT
END_TYPE

(* ---- dfc_moxemm_smu_alm2_4-DFC_MOXEMM_SMU_ALM2_4.st ---- *)
(* --- Interface --- *)
{attribute 'external_name' := 'cmp_rts_DFC_MOXEMM_SMU_ALM2_4'}
TYPE DFC_MOXEMM_SMU_ALM2_4 : STRUCT
		DTC            : UDINT := 16#107E00;
		DFCid          : UINT  := 1233;
		debounceMethod : USINT := NATIVE;
	END_STRUCT
END_TYPE

(* ---- dfc_moxemm_smu_alm2_5-DFC_MOXEMM_SMU_ALM2_5.st ---- *)
(* --- Interface --- *)
{attribute 'external_name' := 'cmp_rts_DFC_MOXEMM_SMU_ALM2_5'}
TYPE DFC_MOXEMM_SMU_ALM2_5 : STRUCT
		DTC            : UDINT := 16#107F00;
		DFCid          : UINT  := 1234;
		debounceMethod : USINT := NATIVE;
	END_STRUCT
END_TYPE

(* ---- dfc_moxemm_smu_alm2_7-DFC_MOXEMM_SMU_ALM2_7.st ---- *)
(* --- Interface --- *)
{attribute 'external_name' := 'cmp_rts_DFC_MOXEMM_SMU_ALM2_7'}
TYPE DFC_MOXEMM_SMU_ALM2_7 : STRUCT
		DTC            : UDINT := 16#108000;
		DFCid          : UINT  := 1235;
		debounceMethod : USINT := NATIVE;
	END_STRUCT
END_TYPE

(* ---- dfc_moxemm_smu_alm2_8-DFC_MOXEMM_SMU_ALM2_8.st ---- *)
(* --- Interface --- *)
{attribute 'external_name' := 'cmp_rts_DFC_MOXEMM_SMU_ALM2_8'}
TYPE DFC_MOXEMM_SMU_ALM2_8 : STRUCT
		DTC            : UDINT := 16#108100;
		DFCid          : UINT  := 1236;
		debounceMethod : USINT := NATIVE;
	END_STRUCT
END_TYPE

(* ---- dfc_moxemm_smu_alm3_1-DFC_MOXEMM_SMU_ALM3_1.st ---- *)
(* --- Interface --- *)
{attribute 'external_name' := 'cmp_rts_DFC_MOXEMM_SMU_ALM3_1'}
TYPE DFC_MOXEMM_SMU_ALM3_1 : STRUCT
		DTC            : UDINT := 16#108800;
		DFCid          : UINT  := 1237;
		debounceMethod : USINT := NATIVE;
	END_STRUCT
END_TYPE

(* ---- dfc_moxemm_smu_alm3_10-DFC_MOXEMM_SMU_ALM3_10.st ---- *)
(* --- Interface --- *)
{attribute 'external_name' := 'cmp_rts_DFC_MOXEMM_SMU_ALM3_10'}
TYPE DFC_MOXEMM_SMU_ALM3_10 : STRUCT
		DTC            : UDINT := 16#108E00;
		DFCid          : UINT  := 1238;
		debounceMethod : USINT := NATIVE;
	END_STRUCT
END_TYPE

(* ---- dfc_moxemm_smu_alm3_11-DFC_MOXEMM_SMU_ALM3_11.st ---- *)
(* --- Interface --- *)
{attribute 'external_name' := 'cmp_rts_DFC_MOXEMM_SMU_ALM3_11'}
TYPE DFC_MOXEMM_SMU_ALM3_11 : STRUCT
		DTC            : UDINT := 16#108F00;
		DFCid          : UINT  := 1239;
		debounceMethod : USINT := NATIVE;
	END_STRUCT
END_TYPE

(* ---- dfc_moxemm_smu_alm3_13-DFC_MOXEMM_SMU_ALM3_13.st ---- *)
(* --- Interface --- *)
{attribute 'external_name' := 'cmp_rts_DFC_MOXEMM_SMU_ALM3_13'}
TYPE DFC_MOXEMM_SMU_ALM3_13 : STRUCT
		DTC            : UDINT := 16#109000;
		DFCid          : UINT  := 1240;
		debounceMethod : USINT := NATIVE;
	END_STRUCT
END_TYPE

(* ---- dfc_moxemm_smu_alm3_14-DFC_MOXEMM_SMU_ALM3_14.st ---- *)
(* --- Interface --- *)
{attribute 'external_name' := 'cmp_rts_DFC_MOXEMM_SMU_ALM3_14'}
TYPE DFC_MOXEMM_SMU_ALM3_14 : STRUCT
		DTC            : UDINT := 16#109100;
		DFCid          : UINT  := 1241;
		debounceMethod : USINT := NATIVE;
	END_STRUCT
END_TYPE

(* ---- dfc_moxemm_smu_alm3_2-DFC_MOXEMM_SMU_ALM3_2.st ---- *)
(* --- Interface --- *)
{attribute 'external_name' := 'cmp_rts_DFC_MOXEMM_SMU_ALM3_2'}
TYPE DFC_MOXEMM_SMU_ALM3_2 : STRUCT
		DTC            : UDINT := 16#108900;
		DFCid          : UINT  := 1242;
		debounceMethod : USINT := NATIVE;
	END_STRUCT
END_TYPE

(* ---- dfc_moxemm_smu_alm3_22-DFC_MOXEMM_SMU_ALM3_22.st ---- *)
(* --- Interface --- *)
{attribute 'external_name' := 'cmp_rts_DFC_MOXEMM_SMU_ALM3_22'}
TYPE DFC_MOXEMM_SMU_ALM3_22 : STRUCT
		DTC            : UDINT := 16#109200;
		DFCid          : UINT  := 1243;
		debounceMethod : USINT := NATIVE;
	END_STRUCT
END_TYPE

(* ---- dfc_moxemm_smu_alm3_23-DFC_MOXEMM_SMU_ALM3_23.st ---- *)
(* --- Interface --- *)
{attribute 'external_name' := 'cmp_rts_DFC_MOXEMM_SMU_ALM3_23'}
TYPE DFC_MOXEMM_SMU_ALM3_23 : STRUCT
		DTC            : UDINT := 16#109300;
		DFCid          : UINT  := 1244;
		debounceMethod : USINT := NATIVE;
	END_STRUCT
END_TYPE

(* ---- dfc_moxemm_smu_alm3_4-DFC_MOXEMM_SMU_ALM3_4.st ---- *)
(* --- Interface --- *)
{attribute 'external_name' := 'cmp_rts_DFC_MOXEMM_SMU_ALM3_4'}
TYPE DFC_MOXEMM_SMU_ALM3_4 : STRUCT
		DTC            : UDINT := 16#108A00;
		DFCid          : UINT  := 1245;
		debounceMethod : USINT := NATIVE;
	END_STRUCT
END_TYPE

(* ---- dfc_moxemm_smu_alm3_5-DFC_MOXEMM_SMU_ALM3_5.st ---- *)
(* --- Interface --- *)
{attribute 'external_name' := 'cmp_rts_DFC_MOXEMM_SMU_ALM3_5'}
TYPE DFC_MOXEMM_SMU_ALM3_5 : STRUCT
		DTC            : UDINT := 16#108B00;
		DFCid          : UINT  := 1246;
		debounceMethod : USINT := NATIVE;
	END_STRUCT
END_TYPE

(* ---- dfc_moxemm_smu_alm3_7-DFC_MOXEMM_SMU_ALM3_7.st ---- *)
(* --- Interface --- *)
{attribute 'external_name' := 'cmp_rts_DFC_MOXEMM_SMU_ALM3_7'}
TYPE DFC_MOXEMM_SMU_ALM3_7 : STRUCT
		DTC            : UDINT := 16#108C00;
		DFCid          : UINT  := 1247;
		debounceMethod : USINT := NATIVE;
	END_STRUCT
END_TYPE

(* ---- dfc_moxemm_smu_alm3_8-DFC_MOXEMM_SMU_ALM3_8.st ---- *)
(* --- Interface --- *)
{attribute 'external_name' := 'cmp_rts_DFC_MOXEMM_SMU_ALM3_8'}
TYPE DFC_MOXEMM_SMU_ALM3_8 : STRUCT
		DTC            : UDINT := 16#108D00;
		DFCid          : UINT  := 1248;
		debounceMethod : USINT := NATIVE;
	END_STRUCT
END_TYPE

(* ---- dfc_moxemm_smu_alm6_0-DFC_MOXEMM_SMU_ALM6_0.st ---- *)
(* --- Interface --- *)
{attribute 'external_name' := 'cmp_rts_DFC_MOXEMM_SMU_ALM6_0'}
TYPE DFC_MOXEMM_SMU_ALM6_0 : STRUCT
		DTC            : UDINT := 16#109400;
		DFCid          : UINT  := 1249;
		debounceMethod : USINT := NATIVE;
	END_STRUCT
END_TYPE

(* ---- dfc_moxemm_smu_alm6_11-DFC_MOXEMM_SMU_ALM6_11.st ---- *)
(* --- Interface --- *)
{attribute 'external_name' := 'cmp_rts_DFC_MOXEMM_SMU_ALM6_11'}
TYPE DFC_MOXEMM_SMU_ALM6_11 : STRUCT
		DTC            : UDINT := 16#109900;
		DFCid          : UINT  := 1250;
		debounceMethod : USINT := NATIVE;
	END_STRUCT
END_TYPE

(* ---- dfc_moxemm_smu_alm6_12-DFC_MOXEMM_SMU_ALM6_12.st ---- *)
(* --- Interface --- *)
{attribute 'external_name' := 'cmp_rts_DFC_MOXEMM_SMU_ALM6_12'}
TYPE DFC_MOXEMM_SMU_ALM6_12 : STRUCT
		DTC            : UDINT := 16#109A00;
		DFCid          : UINT  := 1251;
		debounceMethod : USINT := NATIVE;
	END_STRUCT
END_TYPE

(* ---- dfc_moxemm_smu_alm6_14-DFC_MOXEMM_SMU_ALM6_14.st ---- *)
(* --- Interface --- *)
{attribute 'external_name' := 'cmp_rts_DFC_MOXEMM_SMU_ALM6_14'}
TYPE DFC_MOXEMM_SMU_ALM6_14 : STRUCT
		DTC            : UDINT := 16#109B00;
		DFCid          : UINT  := 1252;
		debounceMethod : USINT := NATIVE;
	END_STRUCT
END_TYPE

(* ---- dfc_moxemm_smu_alm6_15-DFC_MOXEMM_SMU_ALM6_15.st ---- *)
(* --- Interface --- *)
{attribute 'external_name' := 'cmp_rts_DFC_MOXEMM_SMU_ALM6_15'}
TYPE DFC_MOXEMM_SMU_ALM6_15 : STRUCT
		DTC            : UDINT := 16#109C00;
		DFCid          : UINT  := 1253;
		debounceMethod : USINT := NATIVE;
	END_STRUCT
END_TYPE

(* ---- dfc_moxemm_smu_alm6_17-DFC_MOXEMM_SMU_ALM6_17.st ---- *)
(* --- Interface --- *)
{attribute 'external_name' := 'cmp_rts_DFC_MOXEMM_SMU_ALM6_17'}
TYPE DFC_MOXEMM_SMU_ALM6_17 : STRUCT
		DTC            : UDINT := 16#109D00;
		DFCid          : UINT  := 1254;
		debounceMethod : USINT := NATIVE;
	END_STRUCT
END_TYPE

(* ---- dfc_moxemm_smu_alm6_18-DFC_MOXEMM_SMU_ALM6_18.st ---- *)
(* --- Interface --- *)
{attribute 'external_name' := 'cmp_rts_DFC_MOXEMM_SMU_ALM6_18'}
TYPE DFC_MOXEMM_SMU_ALM6_18 : STRUCT
		DTC            : UDINT := 16#109E00;
		DFCid          : UINT  := 1255;
		debounceMethod : USINT := NATIVE;
	END_STRUCT
END_TYPE

(* ---- dfc_moxemm_smu_alm6_2-DFC_MOXEMM_SMU_ALM6_2.st ---- *)
(* --- Interface --- *)
{attribute 'external_name' := 'cmp_rts_DFC_MOXEMM_SMU_ALM6_2'}
TYPE DFC_MOXEMM_SMU_ALM6_2 : STRUCT
		DTC            : UDINT := 16#10D900;
		DFCid          : UINT  := 1256;
		debounceMethod : USINT := NATIVE;
	END_STRUCT
END_TYPE

(* ---- dfc_moxemm_smu_alm6_20-DFC_MOXEMM_SMU_ALM6_20.st ---- *)
(* --- Interface --- *)
{attribute 'external_name' := 'cmp_rts_DFC_MOXEMM_SMU_ALM6_20'}
TYPE DFC_MOXEMM_SMU_ALM6_20 : STRUCT
		DTC            : UDINT := 16#109F00;
		DFCid          : UINT  := 1257;
		debounceMethod : USINT := NATIVE;
	END_STRUCT
END_TYPE

(* ---- dfc_moxemm_smu_alm6_21-DFC_MOXEMM_SMU_ALM6_21.st ---- *)
(* --- Interface --- *)
{attribute 'external_name' := 'cmp_rts_DFC_MOXEMM_SMU_ALM6_21'}
TYPE DFC_MOXEMM_SMU_ALM6_21 : STRUCT
		DTC            : UDINT := 16#10A000;
		DFCid          : UINT  := 1258;
		debounceMethod : USINT := NATIVE;
	END_STRUCT
END_TYPE

(* ---- dfc_moxemm_smu_alm6_25-DFC_MOXEMM_SMU_ALM6_25.st ---- *)
(* --- Interface --- *)
{attribute 'external_name' := 'cmp_rts_DFC_MOXEMM_SMU_ALM6_25'}
TYPE DFC_MOXEMM_SMU_ALM6_25 : STRUCT
		DTC            : UDINT := 16#10A100;
		DFCid          : UINT  := 1259;
		debounceMethod : USINT := NATIVE;
	END_STRUCT
END_TYPE

(* ---- dfc_moxemm_smu_alm6_4-DFC_MOXEMM_SMU_ALM6_4.st ---- *)
(* --- Interface --- *)
{attribute 'external_name' := 'cmp_rts_DFC_MOXEMM_SMU_ALM6_4'}
TYPE DFC_MOXEMM_SMU_ALM6_4 : STRUCT
		DTC            : UDINT := 16#109500;
		DFCid          : UINT  := 1260;
		debounceMethod : USINT := NATIVE;
	END_STRUCT
END_TYPE

(* ---- dfc_moxemm_smu_alm6_5-DFC_MOXEMM_SMU_ALM6_5.st ---- *)
(* --- Interface --- *)
{attribute 'external_name' := 'cmp_rts_DFC_MOXEMM_SMU_ALM6_5'}
TYPE DFC_MOXEMM_SMU_ALM6_5 : STRUCT
		DTC            : UDINT := 16#109600;
		DFCid          : UINT  := 1261;
		debounceMethod : USINT := NATIVE;
	END_STRUCT
END_TYPE

(* ---- dfc_moxemm_smu_alm6_7-DFC_MOXEMM_SMU_ALM6_7.st ---- *)
(* --- Interface --- *)
{attribute 'external_name' := 'cmp_rts_DFC_MOXEMM_SMU_ALM6_7'}
TYPE DFC_MOXEMM_SMU_ALM6_7 : STRUCT
		DTC            : UDINT := 16#109700;
		DFCid          : UINT  := 1262;
		debounceMethod : USINT := NATIVE;
	END_STRUCT
END_TYPE

(* ---- dfc_moxemm_smu_alm6_8-DFC_MOXEMM_SMU_ALM6_8.st ---- *)
(* --- Interface --- *)
{attribute 'external_name' := 'cmp_rts_DFC_MOXEMM_SMU_ALM6_8'}
TYPE DFC_MOXEMM_SMU_ALM6_8 : STRUCT
		DTC            : UDINT := 16#109800;
		DFCid          : UINT  := 1263;
		debounceMethod : USINT := NATIVE;
	END_STRUCT
END_TYPE

(* ---- dfc_moxemm_smu_alm7_1-DFC_MOXEMM_SMU_ALM7_1.st ---- *)
(* --- Interface --- *)
{attribute 'external_name' := 'cmp_rts_DFC_MOXEMM_SMU_ALM7_1'}
TYPE DFC_MOXEMM_SMU_ALM7_1 : STRUCT
		DTC            : UDINT := 16#10A200;
		DFCid          : UINT  := 1264;
		debounceMethod : USINT := NATIVE;
	END_STRUCT
END_TYPE

(* ---- dfc_moxemm_smu_alm7_12-DFC_MOXEMM_SMU_ALM7_12.st ---- *)
(* --- Interface --- *)
{attribute 'external_name' := 'cmp_rts_DFC_MOXEMM_SMU_ALM7_12'}
TYPE DFC_MOXEMM_SMU_ALM7_12 : STRUCT
		DTC            : UDINT := 16#10A400;
		DFCid          : UINT  := 1265;
		debounceMethod : USINT := NATIVE;
	END_STRUCT
END_TYPE

(* ---- dfc_moxemm_smu_alm7_13-DFC_MOXEMM_SMU_ALM7_13.st ---- *)
(* --- Interface --- *)
{attribute 'external_name' := 'cmp_rts_DFC_MOXEMM_SMU_ALM7_13'}
TYPE DFC_MOXEMM_SMU_ALM7_13 : STRUCT
		DTC            : UDINT := 16#10A500;
		DFCid          : UINT  := 1266;
		debounceMethod : USINT := NATIVE;
	END_STRUCT
END_TYPE

(* ---- dfc_moxemm_smu_alm7_14-DFC_MOXEMM_SMU_ALM7_14.st ---- *)
(* --- Interface --- *)
{attribute 'external_name' := 'cmp_rts_DFC_MOXEMM_SMU_ALM7_14'}
TYPE DFC_MOXEMM_SMU_ALM7_14 : STRUCT
		DTC            : UDINT := 16#10A600;
		DFCid          : UINT  := 1267;
		debounceMethod : USINT := NATIVE;
	END_STRUCT
END_TYPE

(* ---- dfc_moxemm_smu_alm7_15-DFC_MOXEMM_SMU_ALM7_15.st ---- *)
(* --- Interface --- *)
{attribute 'external_name' := 'cmp_rts_DFC_MOXEMM_SMU_ALM7_15'}
TYPE DFC_MOXEMM_SMU_ALM7_15 : STRUCT
		DTC            : UDINT := 16#10A700;
		DFCid          : UINT  := 1268;
		debounceMethod : USINT := NATIVE;
	END_STRUCT
END_TYPE

(* ---- dfc_moxemm_smu_alm7_16-DFC_MOXEMM_SMU_ALM7_16.st ---- *)
(* --- Interface --- *)
{attribute 'external_name' := 'cmp_rts_DFC_MOXEMM_SMU_ALM7_16'}
TYPE DFC_MOXEMM_SMU_ALM7_16 : STRUCT
		DTC            : UDINT := 16#10A800;
		DFCid          : UINT  := 1269;
		debounceMethod : USINT := NATIVE;
	END_STRUCT
END_TYPE

(* ---- dfc_moxemm_smu_alm7_17-DFC_MOXEMM_SMU_ALM7_17.st ---- *)
(* --- Interface --- *)
{attribute 'external_name' := 'cmp_rts_DFC_MOXEMM_SMU_ALM7_17'}
TYPE DFC_MOXEMM_SMU_ALM7_17 : STRUCT
		DTC            : UDINT := 16#10A900;
		DFCid          : UINT  := 1270;
		debounceMethod : USINT := NATIVE;
	END_STRUCT
END_TYPE

(* ---- dfc_moxemm_smu_alm7_2-DFC_MOXEMM_SMU_ALM7_2.st ---- *)
(* --- Interface --- *)
{attribute 'external_name' := 'cmp_rts_DFC_MOXEMM_SMU_ALM7_2'}
TYPE DFC_MOXEMM_SMU_ALM7_2 : STRUCT
		DTC            : UDINT := 16#10A300;
		DFCid          : UINT  := 1271;
		debounceMethod : USINT := NATIVE;
	END_STRUCT
END_TYPE

(* ---- dfc_moxemm_smu_alm7_20-DFC_MOXEMM_SMU_ALM7_20.st ---- *)
(* --- Interface --- *)
{attribute 'external_name' := 'cmp_rts_DFC_MOXEMM_SMU_ALM7_20'}
TYPE DFC_MOXEMM_SMU_ALM7_20 : STRUCT
		DTC            : UDINT := 16#10AA00;
		DFCid          : UINT  := 1272;
		debounceMethod : USINT := NATIVE;
	END_STRUCT
END_TYPE

(* ---- dfc_moxemm_smu_alm7_25-DFC_MOXEMM_SMU_ALM7_25.st ---- *)
(* --- Interface --- *)
{attribute 'external_name' := 'cmp_rts_DFC_MOXEMM_SMU_ALM7_25'}
TYPE DFC_MOXEMM_SMU_ALM7_25 : STRUCT
		DTC            : UDINT := 16#10AB00;
		DFCid          : UINT  := 1273;
		debounceMethod : USINT := NATIVE;
	END_STRUCT
END_TYPE

(* ---- dfc_moxemm_smu_alm7_26-DFC_MOXEMM_SMU_ALM7_26.st ---- *)
(* --- Interface --- *)
{attribute 'external_name' := 'cmp_rts_DFC_MOXEMM_SMU_ALM7_26'}
TYPE DFC_MOXEMM_SMU_ALM7_26 : STRUCT
		DTC            : UDINT := 16#10AC00;
		DFCid          : UINT  := 1274;
		debounceMethod : USINT := NATIVE;
	END_STRUCT
END_TYPE

(* ---- dfc_moxemm_smu_alm7_28-DFC_MOXEMM_SMU_ALM7_28.st ---- *)
(* --- Interface --- *)
{attribute 'external_name' := 'cmp_rts_DFC_MOXEMM_SMU_ALM7_28'}
TYPE DFC_MOXEMM_SMU_ALM7_28 : STRUCT
		DTC            : UDINT := 16#10AD00;
		DFCid          : UINT  := 1275;
		debounceMethod : USINT := NATIVE;
	END_STRUCT
END_TYPE

(* ---- dfc_moxemm_smu_alm7_29-DFC_MOXEMM_SMU_ALM7_29.st ---- *)
(* --- Interface --- *)
{attribute 'external_name' := 'cmp_rts_DFC_MOXEMM_SMU_ALM7_29'}
TYPE DFC_MOXEMM_SMU_ALM7_29 : STRUCT
		DTC            : UDINT := 16#10AE00;
		DFCid          : UINT  := 1276;
		debounceMethod : USINT := NATIVE;
	END_STRUCT
END_TYPE

(* ---- dfc_moxemm_smu_alm7_30-DFC_MOXEMM_SMU_ALM7_30.st ---- *)
(* --- Interface --- *)
{attribute 'external_name' := 'cmp_rts_DFC_MOXEMM_SMU_ALM7_30'}
TYPE DFC_MOXEMM_SMU_ALM7_30 : STRUCT
		DTC            : UDINT := 16#10AF00;
		DFCid          : UINT  := 1277;
		debounceMethod : USINT := NATIVE;
	END_STRUCT
END_TYPE

(* ---- dfc_moxemm_smu_alm7_31-DFC_MOXEMM_SMU_ALM7_31.st ---- *)
(* --- Interface --- *)
{attribute 'external_name' := 'cmp_rts_DFC_MOXEMM_SMU_ALM7_31'}
TYPE DFC_MOXEMM_SMU_ALM7_31 : STRUCT
		DTC            : UDINT := 16#10B000;
		DFCid          : UINT  := 1278;
		debounceMethod : USINT := NATIVE;
	END_STRUCT
END_TYPE

(* ---- dfc_moxemm_smu_alm8_0-DFC_MOXEMM_SMU_ALM8_0.st ---- *)
(* --- Interface --- *)
{attribute 'external_name' := 'cmp_rts_DFC_MOXEMM_SMU_ALM8_0'}
TYPE DFC_MOXEMM_SMU_ALM8_0 : STRUCT
		DTC            : UDINT := 16#10B100;
		DFCid          : UINT  := 1279;
		debounceMethod : USINT := NATIVE;
	END_STRUCT
END_TYPE

(* ---- dfc_moxemm_smu_alm8_1-DFC_MOXEMM_SMU_ALM8_1.st ---- *)
(* --- Interface --- *)
{attribute 'external_name' := 'cmp_rts_DFC_MOXEMM_SMU_ALM8_1'}
TYPE DFC_MOXEMM_SMU_ALM8_1 : STRUCT
		DTC            : UDINT := 16#10B200;
		DFCid          : UINT  := 1280;
		debounceMethod : USINT := NATIVE;
	END_STRUCT
END_TYPE

(* ---- dfc_moxemm_smu_alm8_10-DFC_MOXEMM_SMU_ALM8_10.st ---- *)
(* --- Interface --- *)
{attribute 'external_name' := 'cmp_rts_DFC_MOXEMM_SMU_ALM8_10'}
TYPE DFC_MOXEMM_SMU_ALM8_10 : STRUCT
		DTC            : UDINT := 16#10B600;
		DFCid          : UINT  := 1281;
		debounceMethod : USINT := NATIVE;
	END_STRUCT
END_TYPE

(* ---- dfc_moxemm_smu_alm8_11-DFC_MOXEMM_SMU_ALM8_11.st ---- *)
(* --- Interface --- *)
{attribute 'external_name' := 'cmp_rts_DFC_MOXEMM_SMU_ALM8_11'}
TYPE DFC_MOXEMM_SMU_ALM8_11 : STRUCT
		DTC            : UDINT := 16#10B700;
		DFCid          : UINT  := 1282;
		debounceMethod : USINT := NATIVE;
	END_STRUCT
END_TYPE

(* ---- dfc_moxemm_smu_alm8_12-DFC_MOXEMM_SMU_ALM8_12.st ---- *)
(* --- Interface --- *)
{attribute 'external_name' := 'cmp_rts_DFC_MOXEMM_SMU_ALM8_12'}
TYPE DFC_MOXEMM_SMU_ALM8_12 : STRUCT
		DTC            : UDINT := 16#10B800;
		DFCid          : UINT  := 1283;
		debounceMethod : USINT := NATIVE;
	END_STRUCT
END_TYPE

(* ---- dfc_moxemm_smu_alm8_13-DFC_MOXEMM_SMU_ALM8_13.st ---- *)
(* --- Interface --- *)
{attribute 'external_name' := 'cmp_rts_DFC_MOXEMM_SMU_ALM8_13'}
TYPE DFC_MOXEMM_SMU_ALM8_13 : STRUCT
		DTC            : UDINT := 16#10B900;
		DFCid          : UINT  := 1284;
		debounceMethod : USINT := NATIVE;
	END_STRUCT
END_TYPE

(* ---- dfc_moxemm_smu_alm8_16-DFC_MOXEMM_SMU_ALM8_16.st ---- *)
(* --- Interface --- *)
{attribute 'external_name' := 'cmp_rts_DFC_MOXEMM_SMU_ALM8_16'}
TYPE DFC_MOXEMM_SMU_ALM8_16 : STRUCT
		DTC            : UDINT := 16#10BA00;
		DFCid          : UINT  := 1285;
		debounceMethod : USINT := NATIVE;
	END_STRUCT
END_TYPE

(* ---- dfc_moxemm_smu_alm8_18-DFC_MOXEMM_SMU_ALM8_18.st ---- *)
(* --- Interface --- *)
{attribute 'external_name' := 'cmp_rts_DFC_MOXEMM_SMU_ALM8_18'}
TYPE DFC_MOXEMM_SMU_ALM8_18 : STRUCT
		DTC            : UDINT := 16#10BB00;
		DFCid          : UINT  := 1286;
		debounceMethod : USINT := NATIVE;
	END_STRUCT
END_TYPE

(* ---- dfc_moxemm_smu_alm8_2-DFC_MOXEMM_SMU_ALM8_2.st ---- *)
(* --- Interface --- *)
{attribute 'external_name' := 'cmp_rts_DFC_MOXEMM_SMU_ALM8_2'}
TYPE DFC_MOXEMM_SMU_ALM8_2 : STRUCT
		DTC            : UDINT := 16#10B300;
		DFCid          : UINT  := 1287;
		debounceMethod : USINT := NATIVE;
	END_STRUCT
END_TYPE

(* ---- dfc_moxemm_smu_alm8_3-DFC_MOXEMM_SMU_ALM8_3.st ---- *)
(* --- Interface --- *)
{attribute 'external_name' := 'cmp_rts_DFC_MOXEMM_SMU_ALM8_3'}
TYPE DFC_MOXEMM_SMU_ALM8_3 : STRUCT
		DTC            : UDINT := 16#10B400;
		DFCid          : UINT  := 1288;
		debounceMethod : USINT := NATIVE;
	END_STRUCT
END_TYPE

(* ---- dfc_moxemm_smu_alm8_30-DFC_MOXEMM_SMU_ALM8_30.st ---- *)
(* --- Interface --- *)
{attribute 'external_name' := 'cmp_rts_DFC_MOXEMM_SMU_ALM8_30'}
TYPE DFC_MOXEMM_SMU_ALM8_30 : STRUCT
		DTC            : UDINT := 16#10BC00;
		DFCid          : UINT  := 1289;
		debounceMethod : USINT := NATIVE;
	END_STRUCT
END_TYPE

(* ---- dfc_moxemm_smu_alm8_31-DFC_MOXEMM_SMU_ALM8_31.st ---- *)
(* --- Interface --- *)
{attribute 'external_name' := 'cmp_rts_DFC_MOXEMM_SMU_ALM8_31'}
TYPE DFC_MOXEMM_SMU_ALM8_31 : STRUCT
		DTC            : UDINT := 16#10BD00;
		DFCid          : UINT  := 1290;
		debounceMethod : USINT := NATIVE;
	END_STRUCT
END_TYPE

(* ---- dfc_moxemm_smu_alm8_4-DFC_MOXEMM_SMU_ALM8_4.st ---- *)
(* --- Interface --- *)
{attribute 'external_name' := 'cmp_rts_DFC_MOXEMM_SMU_ALM8_4'}
TYPE DFC_MOXEMM_SMU_ALM8_4 : STRUCT
		DTC            : UDINT := 16#10B500;
		DFCid          : UINT  := 1291;
		debounceMethod : USINT := NATIVE;
	END_STRUCT
END_TYPE

(* ---- dfc_moxemm_smu_alm9_0-DFC_MOXEMM_SMU_ALM9_0.st ---- *)
(* --- Interface --- *)
{attribute 'external_name' := 'cmp_rts_DFC_MOXEMM_SMU_ALM9_0'}
TYPE DFC_MOXEMM_SMU_ALM9_0 : STRUCT
		DTC            : UDINT := 16#10BE00;
		DFCid          : UINT  := 1292;
		debounceMethod : USINT := NATIVE;
	END_STRUCT
END_TYPE

(* ---- dfc_moxemm_smu_alm9_1-DFC_MOXEMM_SMU_ALM9_1.st ---- *)
(* --- Interface --- *)
{attribute 'external_name' := 'cmp_rts_DFC_MOXEMM_SMU_ALM9_1'}
TYPE DFC_MOXEMM_SMU_ALM9_1 : STRUCT
		DTC            : UDINT := 16#10BF00;
		DFCid          : UINT  := 1293;
		debounceMethod : USINT := NATIVE;
	END_STRUCT
END_TYPE

(* ---- dfc_moxemm_smu_alm9_15-DFC_MOXEMM_SMU_ALM9_15.st ---- *)
(* --- Interface --- *)
{attribute 'external_name' := 'cmp_rts_DFC_MOXEMM_SMU_ALM9_15'}
TYPE DFC_MOXEMM_SMU_ALM9_15 : STRUCT
		DTC            : UDINT := 16#10C100;
		DFCid          : UINT  := 1294;
		debounceMethod : USINT := NATIVE;
	END_STRUCT
END_TYPE

(* ---- dfc_moxemm_smu_alm9_3-DFC_MOXEMM_SMU_ALM9_3.st ---- *)
(* --- Interface --- *)
{attribute 'external_name' := 'cmp_rts_DFC_MOXEMM_SMU_ALM9_3'}
TYPE DFC_MOXEMM_SMU_ALM9_3 : STRUCT
		DTC            : UDINT := 16#10C000;
		DFCid          : UINT  := 1295;
		debounceMethod : USINT := NATIVE;
	END_STRUCT
END_TYPE

(* ---- dfc_moxemmhwltlbist-DFC_MoXEMMHwLTLBIST.st ---- *)
(* --- Interface --- *)
{attribute 'external_name' := 'cmp_rts_DFC_MoXEMMHwLTLBIST'}
TYPE DFC_MoXEMMHwLTLBIST : STRUCT
		DTC : UDINT := 16#10D000;
	END_STRUCT
END_TYPE

(* ---- dfc_moxemmhwltmbist-DFC_MoXEMMHwLTMBIST.st ---- *)
(* --- Interface --- *)
{attribute 'external_name' := 'cmp_rts_DFC_MoXEMMHwLTMBIST'}
TYPE DFC_MoXEMMHwLTMBIST : STRUCT
		DTC : UDINT := 16#10D100;
	END_STRUCT
END_TYPE

(* ---- dfc_moxemmhwltmcufw-DFC_MoXEMMHwLTMCUFW.st ---- *)
(* --- Interface --- *)
{attribute 'external_name' := 'cmp_rts_DFC_MoXEMMHwLTMCUFW'}
TYPE DFC_MoXEMMHwLTMCUFW : STRUCT
		DTC            : UDINT := 16#10D200;
		DFCid          : UINT  := 1299;
		debounceMethod : USINT := NATIVE;
	END_STRUCT
END_TYPE

(* ---- dfc_moxemmhwltmonbist-DFC_MoXEMMHwLTMonBIST.st ---- *)
(* --- Interface --- *)
{attribute 'external_name' := 'cmp_rts_DFC_MoXEMMHwLTMonBIST'}
TYPE DFC_MoXEMMHwLTMonBIST : STRUCT
		DTC            : UDINT := 16#10D300;
		DFCid          : UINT  := 1300;
		debounceMethod : USINT := NATIVE;
	END_STRUCT
END_TYPE

(* ---- dfc_moxemmhwltregmontest-DFC_MoXEMMHwLTRegMonTest.st ---- *)
(* --- Interface --- *)
{attribute 'external_name' := 'cmp_rts_DFC_MoXEMMHwLTRegMonTest'}
TYPE DFC_MoXEMMHwLTRegMonTest : STRUCT
		DTC            : UDINT := 16#10D400;
		DFCid          : UINT  := 1301;
		debounceMethod : USINT := NATIVE;
	END_STRUCT
END_TYPE

(* ---- dfc_moxemmhwltstbysmualvtest-DFC_MoXEMMHwLTStbySMUAlvTest.st ---- *)
(* --- Interface --- *)
{attribute 'external_name' := 'cmp_rts_DFC_MoXEMMHwLTStbySMUAlvTest'}
TYPE DFC_MoXEMMHwLTStbySMUAlvTest : STRUCT
		DTC            : UDINT := 16#10D500;
		DFCid          : UINT  := 1302;
		debounceMethod : USINT := NATIVE;
	END_STRUCT
END_TYPE

(* ---- dfc_moxemmhwlttempsens-DFC_MoXEMMHwLTTempSens.st ---- *)
(* --- Interface --- *)
{attribute 'external_name' := 'cmp_rts_DFC_MoXEMMHwLTTempSens'}
TYPE DFC_MoXEMMHwLTTempSens : STRUCT
		DTC            : UDINT := 16#10D600;
		DFCid          : UINT  := 1303;
		debounceMethod : USINT := NATIVE;
	END_STRUCT
END_TYPE

(* ---- dfc_moxemmhwltucbcfg-DFC_MoXEMMHwLTUCBCfg.st ---- *)
(* --- Interface --- *)
{attribute 'external_name' := 'cmp_rts_DFC_MoXEMMHwLTUCBCfg'}
TYPE DFC_MoXEMMHwLTUCBCfg : STRUCT
		DTC            : UDINT := 16#10D700;
		DFCid          : UINT  := 1304;
		debounceMethod : USINT := NATIVE;
	END_STRUCT
END_TYPE

(* ---- dfc_mrlyol-DFC_MRlyOL.st ---- *)
(* --- Interface --- *)
{attribute 'external_name' := 'cmp_rts_DFC_MRlyOL'}
TYPE DFC_MRlyOL : STRUCT
		DTC : UDINT := 16#104900;
	END_STRUCT
END_TYPE

(* ---- dfc_mrlyscb-DFC_MRlySCB.st ---- *)
(* --- Interface --- *)
{attribute 'external_name' := 'cmp_rts_DFC_MRlySCB'}
TYPE DFC_MRlySCB : STRUCT
		DTC : UDINT := 16#104A00;
	END_STRUCT
END_TYPE

(* ---- dfc_mrlyscg-DFC_MRlySCG.st ---- *)
(* --- Interface --- *)
{attribute 'external_name' := 'cmp_rts_DFC_MRlySCG'}
TYPE DFC_MRlySCG : STRUCT
		DTC : UDINT := 16#104B00;
	END_STRUCT
END_TYPE

(* ---- dfc_ocwdaabeactv-DFC_OCWDAABEActv.st ---- *)
(* --- Interface --- *)
{attribute 'external_name' := 'cmp_rts_DFC_OCWDAABEActv'}
TYPE DFC_OCWDAABEActv : STRUCT
		DTC            : UDINT := 16#10D800;
		DFCid          : UINT  := 1305;
		debounceMethod : USINT := NATIVE;
	END_STRUCT
END_TYPE

(* ---- dfc_ocwdacom-DFC_OCWDACom.st ---- *)
(* --- Interface --- *)
{attribute 'external_name' := 'cmp_rts_DFC_OCWDACom'}
TYPE DFC_OCWDACom : STRUCT
		DTC            : UDINT := 16#098A00;
		DFCid          : UINT  := 1306;
		debounceMethod : USINT := NATIVE;
	END_STRUCT
END_TYPE

(* ---- dfc_ocwdaerrpin-DFC_OCWDAErrPin.st ---- *)
(* --- Interface --- *)
{attribute 'external_name' := 'cmp_rts_DFC_OCWDAErrPin'}
TYPE DFC_OCWDAErrPin : STRUCT
		DTC            : UDINT := 16#098B00;
		DFCid          : UINT  := 1307;
		debounceMethod : USINT := NATIVE;
	END_STRUCT
END_TYPE

(* ---- dfc_rba_ioextlib_keepalive_drv-DFC_RBA_IOEXTLIB_KEEPALIVE_DRV.st ---- *)
(* --- Interface --- *)
{attribute 'external_name' := 'cmp_rts_DFC_RBA_IOEXTLIB_KEEPALIVE_DRV'}
TYPE DFC_RBA_IOEXTLIB_KEEPALIVE_DRV : STRUCT
		DTC            : UDINT := 16#094300;
		DFCid          : UINT  := 1175;
		debounceMethod : USINT := NO_DEBOUNCE;
	END_STRUCT
END_TYPE

(* ---- dfc_rba_ioextlib_keepalive_ini-DFC_RBA_IOEXTLIB_KEEPALIVE_INI.st ---- *)
(* --- Interface --- *)
{attribute 'external_name' := 'cmp_rts_DFC_RBA_IOEXTLIB_KEEPALIVE_INI'}
TYPE DFC_RBA_IOEXTLIB_KEEPALIVE_INI : STRUCT
		DTC            : UDINT := 16#094400;
		DFCid          : UINT  := 1176;
		debounceMethod : USINT := NO_DEBOUNCE;
	END_STRUCT
END_TYPE

(* ---- dfc_rba_memdiag_memreaderr-DFC_rba_MemDiag_MemReadErr.st ---- *)
(* --- Interface --- *)
{attribute 'external_name' := 'cmp_rts_DFC_rba_MemDiag_MemReadErr'}
TYPE DFC_rba_MemDiag_MemReadErr : STRUCT
		DTC            : UDINT := 16#094700;
		DFCid          : UINT  := 1179;
		debounceMethod : USINT := NO_DEBOUNCE;
	END_STRUCT
END_TYPE

(* ---- dfc_rba_memdiag_memwrerr-DFC_rba_MemDiag_MemWrErr.st ---- *)
(* --- Interface --- *)
{attribute 'external_name' := 'cmp_rts_DFC_rba_MemDiag_MemWrErr'}
TYPE DFC_rba_MemDiag_MemWrErr : STRUCT
		DTC            : UDINT := 16#094800;
		DFCid          : UINT  := 1180;
		debounceMethod : USINT := NO_DEBOUNCE;
	END_STRUCT
END_TYPE

(* ---- dfc_rba_memdiagextd_memreadsngerr-DFC_rba_MemDiagExtd_MemReadSngErr.st ---- *)
(* --- Interface --- *)
{attribute 'external_name' := 'cmp_rts_DFC_rba_MemDiagExtd_MemReadSngErr'}
TYPE DFC_rba_MemDiagExtd_MemReadSngErr : STRUCT
		DTC            : UDINT := 16#103E00;
		DFCid          : UINT  := 1178;
		debounceMethod : USINT := NO_DEBOUNCE;
	END_STRUCT
END_TYPE

(* ---- dfc_rba_mrly_diag_stk_event-DFC_rba_MRly_Diag_Stk_Event.st ---- *)
(* --- Interface --- *)
{attribute 'external_name' := 'cmp_rts_DFC_rba_MRly_Diag_Stk_Event'}
TYPE DFC_rba_MRly_Diag_Stk_Event : STRUCT
		DTC            : UDINT := 16#094600;
		DFCid          : UINT  := 1177;
		debounceMethod : USINT := NO_DEBOUNCE;
	END_STRUCT
END_TYPE

(* ---- dfc_rba_multistacktrace_threshold-DFC_rba_MultiStackTrace_Threshold.st ---- *)
(* --- Interface --- *)
{attribute 'external_name' := 'cmp_rts_DFC_rba_MultiStackTrace_Threshold'}
TYPE DFC_rba_MultiStackTrace_Threshold : STRUCT
		DTC            : UDINT := 16#094900;
		DFCid          : UINT  := 1173;
		debounceMethod : USINT := NO_DEBOUNCE;
	END_STRUCT
END_TYPE

(* ---- dfc_rba_syc_irrswofftrigengrun_event-DFC_rba_SyC_IrrSwOffTrigEngRun_Event.st ---- *)
(* --- Interface --- *)
{attribute 'external_name' := 'cmp_rts_DFC_rba_SyC_IrrSwOffTrigEngRun_Event'}
TYPE DFC_rba_SyC_IrrSwOffTrigEngRun_Event : STRUCT
		DTC            : UDINT := 16#094A00;
		DFCid          : UINT  := 1181;
		debounceMethod : USINT := NO_DEBOUNCE;
	END_STRUCT
END_TYPE

(* ---- dfc_rba_t15_diag_cominvld_event-DFC_rba_T15_Diag_ComInVld_Event.st ---- *)
(* --- Interface --- *)
{attribute 'external_name' := 'cmp_rts_DFC_rba_T15_Diag_ComInVld_Event'}
TYPE DFC_rba_T15_Diag_ComInVld_Event : STRUCT
		DTC            : UDINT := 16#094B00;
		DFCid          : UINT  := 1182;
		debounceMethod : USINT := NO_DEBOUNCE;
	END_STRUCT
END_TYPE

(* ---- dfc_rba_t15_diag_comoff_hwon_event-DFC_rba_T15_Diag_ComOff_HwOn_Event.st ---- *)
(* --- Interface --- *)
{attribute 'external_name' := 'cmp_rts_DFC_rba_T15_Diag_ComOff_HwOn_Event'}
TYPE DFC_rba_T15_Diag_ComOff_HwOn_Event : STRUCT
		DTC            : UDINT := 16#094C00;
		DFCid          : UINT  := 1183;
		debounceMethod : USINT := NO_DEBOUNCE;
	END_STRUCT
END_TYPE

(* ---- dfc_rba_t15_diag_comon_hwoff_event-DFC_rba_T15_Diag_ComOn_HwOff_Event.st ---- *)
(* --- Interface --- *)
{attribute 'external_name' := 'cmp_rts_DFC_rba_T15_Diag_ComOn_HwOff_Event'}
TYPE DFC_rba_T15_Diag_ComOn_HwOff_Event : STRUCT
		DTC            : UDINT := 16#094D00;
		DFCid          : UINT  := 1184;
		debounceMethod : USINT := NO_DEBOUNCE;
	END_STRUCT
END_TYPE

(* ---- dfc_rbr_can_clearipdugroup-DFC_rbr_can_ClearIpduGroup.st ---- *)
(* --- Interface --- *)
{attribute 'external_name' := 'cmp_rts_DFC_rbr_can_ClearIpduGroup'}
TYPE DFC_rbr_can_ClearIpduGroup : STRUCT
		DTC            : UDINT := 16#022C00;
		DFCid          : UINT  := 864;
		debounceMethod : USINT := NO_DEBOUNCE;
	END_STRUCT
END_TYPE

(* ---- dfc_rbr_can_receivesignal-DFC_rbr_can_ReceiveSignal.st ---- *)
(* --- Interface --- *)
{attribute 'external_name' := 'cmp_rts_DFC_rbr_can_ReceiveSignal'}
TYPE DFC_rbr_can_ReceiveSignal : STRUCT
		DTC            : UDINT := 16#022A00;
		DFCid          : UINT  := 865;
		debounceMethod : USINT := NO_DEBOUNCE;
	END_STRUCT
END_TYPE

(* ---- dfc_rbr_can_sendsignal-DFC_rbr_can_SendSignal.st ---- *)
(* --- Interface --- *)
{attribute 'external_name' := 'cmp_rts_DFC_rbr_can_SendSignal'}
TYPE DFC_rbr_can_SendSignal : STRUCT
		DTC            : UDINT := 16#022900;
		DFCid          : UINT  := 866;
		debounceMethod : USINT := NO_DEBOUNCE;
	END_STRUCT
END_TYPE

(* ---- dfc_rbr_can_setipdugroup-DFC_rbr_can_SetIpduGroup.st ---- *)
(* --- Interface --- *)
{attribute 'external_name' := 'cmp_rts_DFC_rbr_can_SetIpduGroup'}
TYPE DFC_rbr_can_SetIpduGroup : STRUCT
		DTC            : UDINT := 16#022B00;
		DFCid          : UINT  := 867;
		debounceMethod : USINT := NO_DEBOUNCE;
	END_STRUCT
END_TYPE

(* ---- dfc_rbr_cangetdataboxnoinit-DFC_rbr_canGetDataboxNoInit.st ---- *)
(* --- Interface --- *)
{attribute 'external_name' := 'cmp_rts_DFC_rbr_canGetDataboxNoInit'}
TYPE DFC_rbr_canGetDataboxNoInit : STRUCT
		DTC            : UDINT := 16#020100;
		DFCid          : UINT  := 825;
		debounceMethod : USINT := NO_DEBOUNCE;
	END_STRUCT
END_TYPE

(* ---- dfc_rbr_cangetdataboxparam-DFC_rbr_canGetDataboxParam.st ---- *)
(* --- Interface --- *)
{attribute 'external_name' := 'cmp_rts_DFC_rbr_canGetDataboxParam'}
TYPE DFC_rbr_canGetDataboxParam : STRUCT
		DTC            : UDINT := 16#020200;
		DFCid          : UINT  := 826;
		debounceMethod : USINT := NO_DEBOUNCE;
	END_STRUCT
END_TYPE

(* ---- dfc_rbr_cangetdatanobuf-DFC_rbr_canGetDataNoBuf.st ---- *)
(* --- Interface --- *)
{attribute 'external_name' := 'cmp_rts_DFC_rbr_canGetDataNoBuf'}
TYPE DFC_rbr_canGetDataNoBuf : STRUCT
		DTC            : UDINT := 16#020300;
		DFCid          : UINT  := 823;
		debounceMethod : USINT := NO_DEBOUNCE;
	END_STRUCT
END_TYPE

(* ---- dfc_rbr_cangetdataparam-DFC_rbr_canGetDataParam.st ---- *)
(* --- Interface --- *)
{attribute 'external_name' := 'cmp_rts_DFC_rbr_canGetDataParam'}
TYPE DFC_rbr_canGetDataParam : STRUCT
		DTC            : UDINT := 16#020400;
		DFCid          : UINT  := 824;
		debounceMethod : USINT := NO_DEBOUNCE;
	END_STRUCT
END_TYPE

(* ---- dfc_rbr_cangetrxbufstatusparam-DFC_rbr_canGetRxBufStatusParam.st ---- *)
(* --- Interface --- *)
{attribute 'external_name' := 'cmp_rts_DFC_rbr_canGetRxBufStatusParam'}
TYPE DFC_rbr_canGetRxBufStatusParam : STRUCT
		DTC            : UDINT := 16#020500;
		DFCid          : UINT  := 827;
		debounceMethod : USINT := NO_DEBOUNCE;
	END_STRUCT
END_TYPE

(* ---- dfc_rbr_cangetstatusparam-DFC_rbr_canGetStatusParam.st ---- *)
(* --- Interface --- *)
{attribute 'external_name' := 'cmp_rts_DFC_rbr_canGetStatusParam'}
TYPE DFC_rbr_canGetStatusParam : STRUCT
		DTC            : UDINT := 16#020600;
		DFCid          : UINT  := 828;
		debounceMethod : USINT := NO_DEBOUNCE;
	END_STRUCT
END_TYPE

(* ---- dfc_rbr_cangettxbufstatusparam-DFC_rbr_canGetTxBufStatusParam.st ---- *)
(* --- Interface --- *)
{attribute 'external_name' := 'cmp_rts_DFC_rbr_canGetTxBufStatusParam'}
TYPE DFC_rbr_canGetTxBufStatusParam : STRUCT
		DTC            : UDINT := 16#020700;
		DFCid          : UINT  := 829;
		debounceMethod : USINT := NO_DEBOUNCE;
	END_STRUCT
END_TYPE

(* ---- dfc_rbr_caninitparam-DFC_rbr_canInitParam.st ---- *)
(* --- Interface --- *)
{attribute 'external_name' := 'cmp_rts_DFC_rbr_canInitParam'}
TYPE DFC_rbr_canInitParam : STRUCT
		DTC            : UDINT := 16#020800;
		DFCid          : UINT  := 830;
		debounceMethod : USINT := NO_DEBOUNCE;
	END_STRUCT
END_TYPE

(* ---- dfc_rbr_caninitrxdataboxoverlap-DFC_rbr_canInitRxDataboxOverlap.st ---- *)
(* --- Interface --- *)
{attribute 'external_name' := 'cmp_rts_DFC_rbr_canInitRxDataboxOverlap'}
TYPE DFC_rbr_canInitRxDataboxOverlap : STRUCT
		DTC            : UDINT := 16#020900;
		DFCid          : UINT  := 831;
		debounceMethod : USINT := NO_DEBOUNCE;
	END_STRUCT
END_TYPE

(* ---- dfc_rbr_caninitrxdataboxparam-DFC_rbr_canInitRxDataboxParam.st ---- *)
(* --- Interface --- *)
{attribute 'external_name' := 'cmp_rts_DFC_rbr_canInitRxDataboxParam'}
TYPE DFC_rbr_canInitRxDataboxParam : STRUCT
		DTC            : UDINT := 16#020A00;
		DFCid          : UINT  := 832;
		debounceMethod : USINT := NO_DEBOUNCE;
	END_STRUCT
END_TYPE

(* ---- dfc_rbr_caninittxdataboxparam-DFC_rbr_canInitTxDataboxParam.st ---- *)
(* --- Interface --- *)
{attribute 'external_name' := 'cmp_rts_DFC_rbr_canInitTxDataboxParam'}
TYPE DFC_rbr_canInitTxDataboxParam : STRUCT
		DTC            : UDINT := 16#020B00;
		DFCid          : UINT  := 833;
		debounceMethod : USINT := NO_DEBOUNCE;
	END_STRUCT
END_TYPE

(* ---- dfc_rbr_canipdugroupcontrol-DFC_rbr_canIpduGroupControl.st ---- *)
(* --- Interface --- *)
{attribute 'external_name' := 'cmp_rts_DFC_rbr_canIpduGroupControl'}
TYPE DFC_rbr_canIpduGroupControl : STRUCT
		DTC            : UDINT := 16#022D00;
		DFCid          : UINT  := 834;
		debounceMethod : USINT := NO_DEBOUNCE;
	END_STRUCT
END_TYPE

(* ---- dfc_rbr_canisdataboxfreenoinit-DFC_rbr_canIsDataboxFreeNoInit.st ---- *)
(* --- Interface --- *)
{attribute 'external_name' := 'cmp_rts_DFC_rbr_canIsDataboxFreeNoInit'}
TYPE DFC_rbr_canIsDataboxFreeNoInit : STRUCT
		DTC            : UDINT := 16#020C00;
		DFCid          : UINT  := 835;
		debounceMethod : USINT := NO_DEBOUNCE;
	END_STRUCT
END_TYPE

(* ---- dfc_rbr_canisdataboxfreeparam-DFC_rbr_canIsDataboxFreeParam.st ---- *)
(* --- Interface --- *)
{attribute 'external_name' := 'cmp_rts_DFC_rbr_canIsDataboxFreeParam'}
TYPE DFC_rbr_canIsDataboxFreeParam : STRUCT
		DTC            : UDINT := 16#020D00;
		DFCid          : UINT  := 836;
		debounceMethod : USINT := NO_DEBOUNCE;
	END_STRUCT
END_TYPE

(* ---- dfc_rbr_canistxemptyparam-DFC_rbr_canIsTxEmptyParam.st ---- *)
(* --- Interface --- *)
{attribute 'external_name' := 'cmp_rts_DFC_rbr_canIsTxEmptyParam'}
TYPE DFC_rbr_canIsTxEmptyParam : STRUCT
		DTC            : UDINT := 16#020E00;
		DFCid          : UINT  := 837;
		debounceMethod : USINT := NO_DEBOUNCE;
	END_STRUCT
END_TYPE

(* ---- dfc_rbr_canregbusoffcallbinvstate-DFC_rbr_canRegBusOffCallbInvState.st ---- *)
(* --- Interface --- *)
{attribute 'external_name' := 'cmp_rts_DFC_rbr_canRegBusOffCallbInvState'}
TYPE DFC_rbr_canRegBusOffCallbInvState : STRUCT
		DTC            : UDINT := 16#020F00;
		DFCid          : UINT  := 838;
		debounceMethod : USINT := NO_DEBOUNCE;
	END_STRUCT
END_TYPE

(* ---- dfc_rbr_canregbusoffcallbparam-DFC_rbr_canRegBusOffCallbParam.st ---- *)
(* --- Interface --- *)
{attribute 'external_name' := 'cmp_rts_DFC_rbr_canRegBusOffCallbParam'}
TYPE DFC_rbr_canRegBusOffCallbParam : STRUCT
		DTC            : UDINT := 16#021000;
		DFCid          : UINT  := 839;
		debounceMethod : USINT := NO_DEBOUNCE;
	END_STRUCT
END_TYPE

(* ---- dfc_rbr_canregrxbufinvstate-DFC_rbr_canRegRxBufInvState.st ---- *)
(* --- Interface --- *)
{attribute 'external_name' := 'cmp_rts_DFC_rbr_canRegRxBufInvState'}
TYPE DFC_rbr_canRegRxBufInvState : STRUCT
		DTC            : UDINT := 16#021100;
		DFCid          : UINT  := 840;
		debounceMethod : USINT := NO_DEBOUNCE;
	END_STRUCT
END_TYPE

(* ---- dfc_rbr_canregrxbufoverlap-DFC_rbr_canRegRxBufOverlap.st ---- *)
(* --- Interface --- *)
{attribute 'external_name' := 'cmp_rts_DFC_rbr_canRegRxBufOverlap'}
TYPE DFC_rbr_canRegRxBufOverlap : STRUCT
		DTC            : UDINT := 16#021200;
		DFCid          : UINT  := 841;
		debounceMethod : USINT := NO_DEBOUNCE;
	END_STRUCT
END_TYPE

(* ---- dfc_rbr_canregrxbufparam-DFC_rbr_canRegRxBufParam.st ---- *)
(* --- Interface --- *)
{attribute 'external_name' := 'cmp_rts_DFC_rbr_canRegRxBufParam'}
TYPE DFC_rbr_canRegRxBufParam : STRUCT
		DTC            : UDINT := 16#021300;
		DFCid          : UINT  := 842;
		debounceMethod : USINT := NO_DEBOUNCE;
	END_STRUCT
END_TYPE

(* ---- dfc_rbr_canregrxcallbinvstate-DFC_rbr_canRegRxCallbInvState.st ---- *)
(* --- Interface --- *)
{attribute 'external_name' := 'cmp_rts_DFC_rbr_canRegRxCallbInvState'}
TYPE DFC_rbr_canRegRxCallbInvState : STRUCT
		DTC            : UDINT := 16#021400;
		DFCid          : UINT  := 843;
		debounceMethod : USINT := NO_DEBOUNCE;
	END_STRUCT
END_TYPE

(* ---- dfc_rbr_canregrxcallbparam-DFC_rbr_canRegRxCallbParam.st ---- *)
(* --- Interface --- *)
{attribute 'external_name' := 'cmp_rts_DFC_rbr_canRegRxCallbParam'}
TYPE DFC_rbr_canRegRxCallbParam : STRUCT
		DTC            : UDINT := 16#021500;
		DFCid          : UINT  := 844;
		debounceMethod : USINT := NO_DEBOUNCE;
	END_STRUCT
END_TYPE

(* ---- dfc_rbr_canregrxdataboxinvnumb-DFC_rbr_canRegRxDataboxInvNumb.st ---- *)
(* --- Interface --- *)
{attribute 'external_name' := 'cmp_rts_DFC_rbr_canRegRxDataboxInvNumb'}
TYPE DFC_rbr_canRegRxDataboxInvNumb : STRUCT
		DTC            : UDINT := 16#021600;
		DFCid          : UINT  := 845;
		debounceMethod : USINT := NO_DEBOUNCE;
	END_STRUCT
END_TYPE

(* ---- dfc_rbr_canregrxdataboxinvstate-DFC_rbr_canRegRxDataboxInvState.st ---- *)
(* --- Interface --- *)
{attribute 'external_name' := 'cmp_rts_DFC_rbr_canRegRxDataboxInvState'}
TYPE DFC_rbr_canRegRxDataboxInvState : STRUCT
		DTC            : UDINT := 16#021700;
		DFCid          : UINT  := 846;
		debounceMethod : USINT := NO_DEBOUNCE;
	END_STRUCT
END_TYPE

(* ---- dfc_rbr_canregrxdataboxoverlap-DFC_rbr_canRegRxDataboxOverlap.st ---- *)
(* --- Interface --- *)
{attribute 'external_name' := 'cmp_rts_DFC_rbr_canRegRxDataboxOverlap'}
TYPE DFC_rbr_canRegRxDataboxOverlap : STRUCT
		DTC            : UDINT := 16#021800;
		DFCid          : UINT  := 847;
		debounceMethod : USINT := NO_DEBOUNCE;
	END_STRUCT
END_TYPE

(* ---- dfc_rbr_canregrxdataboxparam-DFC_rbr_canRegRxDataboxParam.st ---- *)
(* --- Interface --- *)
{attribute 'external_name' := 'cmp_rts_DFC_rbr_canRegRxDataboxParam'}
TYPE DFC_rbr_canRegRxDataboxParam : STRUCT
		DTC            : UDINT := 16#021900;
		DFCid          : UINT  := 848;
		debounceMethod : USINT := NO_DEBOUNCE;
	END_STRUCT
END_TYPE

(* ---- dfc_rbr_canregtxbufinvstate-DFC_rbr_canRegTxBufInvState.st ---- *)
(* --- Interface --- *)
{attribute 'external_name' := 'cmp_rts_DFC_rbr_canRegTxBufInvState'}
TYPE DFC_rbr_canRegTxBufInvState : STRUCT
		DTC            : UDINT := 16#021A00;
		DFCid          : UINT  := 849;
		debounceMethod : USINT := NO_DEBOUNCE;
	END_STRUCT
END_TYPE

(* ---- dfc_rbr_canregtxbufoverlap-DFC_rbr_canRegTxBufOverlap.st ---- *)
(* --- Interface --- *)
{attribute 'external_name' := 'cmp_rts_DFC_rbr_canRegTxBufOverlap'}
TYPE DFC_rbr_canRegTxBufOverlap : STRUCT
		DTC            : UDINT := 16#021B00;
		DFCid          : UINT  := 850;
		debounceMethod : USINT := NO_DEBOUNCE;
	END_STRUCT
END_TYPE

(* ---- dfc_rbr_canregtxbufparam-DFC_rbr_canRegTxBufParam.st ---- *)
(* --- Interface --- *)
{attribute 'external_name' := 'cmp_rts_DFC_rbr_canRegTxBufParam'}
TYPE DFC_rbr_canRegTxBufParam : STRUCT
		DTC            : UDINT := 16#021C00;
		DFCid          : UINT  := 851;
		debounceMethod : USINT := NO_DEBOUNCE;
	END_STRUCT
END_TYPE

(* ---- dfc_rbr_canregtxdataboxinvnumb-DFC_rbr_canRegTxDataboxInvNumb.st ---- *)
(* --- Interface --- *)
{attribute 'external_name' := 'cmp_rts_DFC_rbr_canRegTxDataboxInvNumb'}
TYPE DFC_rbr_canRegTxDataboxInvNumb : STRUCT
		DTC            : UDINT := 16#021D00;
		DFCid          : UINT  := 852;
		debounceMethod : USINT := NO_DEBOUNCE;
	END_STRUCT
END_TYPE

(* ---- dfc_rbr_canregtxdataboxinvstate-DFC_rbr_canRegTxDataboxInvState.st ---- *)
(* --- Interface --- *)
{attribute 'external_name' := 'cmp_rts_DFC_rbr_canRegTxDataboxInvState'}
TYPE DFC_rbr_canRegTxDataboxInvState : STRUCT
		DTC            : UDINT := 16#021E00;
		DFCid          : UINT  := 853;
		debounceMethod : USINT := NO_DEBOUNCE;
	END_STRUCT
END_TYPE

(* ---- dfc_rbr_canregtxdataboxoverlap-DFC_rbr_canRegTxDataboxOverlap.st ---- *)
(* --- Interface --- *)
{attribute 'external_name' := 'cmp_rts_DFC_rbr_canRegTxDataboxOverlap'}
TYPE DFC_rbr_canRegTxDataboxOverlap : STRUCT
		DTC            : UDINT := 16#021F00;
		DFCid          : UINT  := 854;
		debounceMethod : USINT := NO_DEBOUNCE;
	END_STRUCT
END_TYPE

(* ---- dfc_rbr_canregtxdataboxparam-DFC_rbr_canRegTxDataboxParam.st ---- *)
(* --- Interface --- *)
{attribute 'external_name' := 'cmp_rts_DFC_rbr_canRegTxDataboxParam'}
TYPE DFC_rbr_canRegTxDataboxParam : STRUCT
		DTC            : UDINT := 16#022000;
		DFCid          : UINT  := 855;
		debounceMethod : USINT := NO_DEBOUNCE;
	END_STRUCT
END_TYPE

(* ---- dfc_rbr_canresettxbufparam-DFC_rbr_canResetTxBufParam.st ---- *)
(* --- Interface --- *)
{attribute 'external_name' := 'cmp_rts_DFC_rbr_canResetTxBufParam'}
TYPE DFC_rbr_canResetTxBufParam : STRUCT
		DTC            : UDINT := 16#022100;
		DFCid          : UINT  := 856;
		debounceMethod : USINT := NO_DEBOUNCE;
	END_STRUCT
END_TYPE

(* ---- dfc_rbr_cansenddataboxnoinit-DFC_rbr_canSendDataboxNoInit.st ---- *)
(* --- Interface --- *)
{attribute 'external_name' := 'cmp_rts_DFC_rbr_canSendDataboxNoInit'}
TYPE DFC_rbr_canSendDataboxNoInit : STRUCT
		DTC            : UDINT := 16#022200;
		DFCid          : UINT  := 859;
		debounceMethod : USINT := NO_DEBOUNCE;
	END_STRUCT
END_TYPE

(* ---- dfc_rbr_cansenddataboxparam-DFC_rbr_canSendDataboxParam.st ---- *)
(* --- Interface --- *)
{attribute 'external_name' := 'cmp_rts_DFC_rbr_canSendDataboxParam'}
TYPE DFC_rbr_canSendDataboxParam : STRUCT
		DTC            : UDINT := 16#022300;
		DFCid          : UINT  := 860;
		debounceMethod : USINT := NO_DEBOUNCE;
	END_STRUCT
END_TYPE

(* ---- dfc_rbr_cansenddatabufovfl-DFC_rbr_canSendDataBufOvfl.st ---- *)
(* --- Interface --- *)
{attribute 'external_name' := 'cmp_rts_DFC_rbr_canSendDataBufOvfl'}
TYPE DFC_rbr_canSendDataBufOvfl : STRUCT
		DTC            : UDINT := 16#022400;
		DFCid          : UINT  := 857;
		debounceMethod : USINT := NO_DEBOUNCE;
	END_STRUCT
END_TYPE

(* ---- dfc_rbr_cansenddataparam-DFC_rbr_canSendDataParam.st ---- *)
(* --- Interface --- *)
{attribute 'external_name' := 'cmp_rts_DFC_rbr_canSendDataParam'}
TYPE DFC_rbr_canSendDataParam : STRUCT
		DTC            : UDINT := 16#022500;
		DFCid          : UINT  := 858;
		debounceMethod : USINT := NO_DEBOUNCE;
	END_STRUCT
END_TYPE

(* ---- dfc_rbr_cansettxcycleparam-DFC_rbr_canSetTxCycleParam.st ---- *)
(* --- Interface --- *)
{attribute 'external_name' := 'cmp_rts_DFC_rbr_canSetTxCycleParam'}
TYPE DFC_rbr_canSetTxCycleParam : STRUCT
		DTC            : UDINT := 16#022600;
		DFCid          : UINT  := 861;
		debounceMethod : USINT := NO_DEBOUNCE;
	END_STRUCT
END_TYPE

(* ---- dfc_rbr_canstartparam-DFC_rbr_canStartParam.st ---- *)
(* --- Interface --- *)
{attribute 'external_name' := 'cmp_rts_DFC_rbr_canStartParam'}
TYPE DFC_rbr_canStartParam : STRUCT
		DTC            : UDINT := 16#022700;
		DFCid          : UINT  := 862;
		debounceMethod : USINT := NO_DEBOUNCE;
	END_STRUCT
END_TYPE

(* ---- dfc_rbr_canstopparam-DFC_rbr_canStopParam.st ---- *)
(* --- Interface --- *)
{attribute 'external_name' := 'cmp_rts_DFC_rbr_canStopParam'}
TYPE DFC_rbr_canStopParam : STRUCT
		DTC            : UDINT := 16#022800;
		DFCid          : UINT  := 863;
		debounceMethod : USINT := NO_DEBOUNCE;
	END_STRUCT
END_TYPE

(* ---- dfc_rbr_dsmdeldtcj1939-DFC_rbr_dsmDelDTCJ1939.st ---- *)
(* --- Interface --- *)
{attribute 'external_name' := 'cmp_rts_DFC_rbr_dsmDelDTCJ1939'}
TYPE DFC_rbr_dsmDelDTCJ1939 : STRUCT
		DTC            : UDINT := 16#070400;
		DFCid          : UINT  := 869;
		debounceMethod : USINT := NO_DEBOUNCE;
	END_STRUCT
END_TYPE

(* ---- dfc_rbr_dsmdelerrors-DFC_rbr_dsmDelErrors.st ---- *)
(* --- Interface --- *)
{attribute 'external_name' := 'cmp_rts_DFC_rbr_dsmDelErrors'}
TYPE DFC_rbr_dsmDelErrors : STRUCT
		DTC            : UDINT := 16#070700;
		DFCid          : UINT  := 870;
		debounceMethod : USINT := NO_DEBOUNCE;
	END_STRUCT
END_TYPE

(* ---- dfc_rbr_dsmdtcj1939-DFC_rbr_dsmDTCJ1939.st ---- *)
(* --- Interface --- *)
{attribute 'external_name' := 'cmp_rts_DFC_rbr_dsmDTCJ1939'}
TYPE DFC_rbr_dsmDTCJ1939 : STRUCT
		DTC            : UDINT := 16#071000;
		DFCid          : UINT  := 868;
		debounceMethod : USINT := NO_DEBOUNCE;
	END_STRUCT
END_TYPE

(* ---- dfc_rbr_dsmgetdfcstatus-DFC_rbr_dsmgetDFCStatus.st ---- *)
(* --- Interface --- *)
{attribute 'external_name' := 'cmp_rts_DFC_rbr_dsmgetDFCStatus'}
TYPE DFC_rbr_dsmgetDFCStatus : STRUCT
		DTC            : UDINT := 16#071100;
		DFCid          : UINT  := 880;
		debounceMethod : USINT := NO_DEBOUNCE;
	END_STRUCT
END_TYPE

(* ---- dfc_rbr_dsmgetdfes-DFC_rbr_dsmGetDFES.st ---- *)
(* --- Interface --- *)
{attribute 'external_name' := 'cmp_rts_DFC_rbr_dsmGetDFES'}
TYPE DFC_rbr_dsmGetDFES : STRUCT
		DTC            : UDINT := 16#070500;
		DFCid          : UINT  := 871;
		debounceMethod : USINT := NO_DEBOUNCE;
	END_STRUCT
END_TYPE

(* ---- dfc_rbr_dsmgetdtcj1939-DFC_rbr_dsmGetDTCJ1939.st ---- *)
(* --- Interface --- *)
{attribute 'external_name' := 'cmp_rts_DFC_rbr_dsmGetDTCJ1939'}
TYPE DFC_rbr_dsmGetDTCJ1939 : STRUCT
		DTC            : UDINT := 16#070300;
		DFCid          : UINT  := 872;
		debounceMethod : USINT := NO_DEBOUNCE;
	END_STRUCT
END_TYPE

(* ---- dfc_rbr_dsmgeterrors-DFC_rbr_dsmGetErrors.st ---- *)
(* --- Interface --- *)
{attribute 'external_name' := 'cmp_rts_DFC_rbr_dsmGetErrors'}
TYPE DFC_rbr_dsmGetErrors : STRUCT
		DTC            : UDINT := 16#070100;
		DFCid          : UINT  := 873;
		debounceMethod : USINT := NO_DEBOUNCE;
	END_STRUCT
END_TYPE

(* ---- dfc_rbr_dsmgetnumerrors-DFC_rbr_dsmGetNumErrors.st ---- *)
(* --- Interface --- *)
{attribute 'external_name' := 'cmp_rts_DFC_rbr_dsmGetNumErrors'}
TYPE DFC_rbr_dsmGetNumErrors : STRUCT
		DTC            : UDINT := 16#070200;
		DFCid          : UINT  := 874;
		debounceMethod : USINT := NO_DEBOUNCE;
	END_STRUCT
END_TYPE

(* ---- dfc_rbr_dsminitqueueoverflow-DFC_rbr_dsmInitQueueOverflow.st ---- *)
(* --- Interface --- *)
{attribute 'external_name' := 'cmp_rts_DFC_rbr_dsmInitQueueOverflow'}
TYPE DFC_rbr_dsmInitQueueOverflow : STRUCT
		DTC            : UDINT := 16#071400;
		DFCid          : UINT  := 875;
		debounceMethod : USINT := NO_DEBOUNCE;
	END_STRUCT
END_TYPE

(* ---- dfc_rbr_dsmnumdtcj1939-DFC_rbr_dsmNumDTCJ1939.st ---- *)
(* --- Interface --- *)
{attribute 'external_name' := 'cmp_rts_DFC_rbr_dsmNumDTCJ1939'}
TYPE DFC_rbr_dsmNumDTCJ1939 : STRUCT
		DTC            : UDINT := 16#071300;
		DFCid          : UINT  := 876;
		debounceMethod : USINT := NO_DEBOUNCE;
	END_STRUCT
END_TYPE

(* ---- dfc_rbr_dsmtesterror-DFC_rbr_dsmTesterror.st ---- *)
(* --- Interface --- *)
{attribute 'external_name' := 'cmp_rts_DFC_rbr_dsmTesterror'}
TYPE DFC_rbr_dsmTesterror : STRUCT
		DTC            : UDINT := 16#070600;
		DFCid          : UINT  := 877;
		debounceMethod : USINT := NO_DEBOUNCE;
	END_STRUCT
END_TYPE

(* ---- dfc_rbr_dsmtesterrordfc-DFC_rbr_dsmtestErrorDFC.st ---- *)
(* --- Interface --- *)
{attribute 'external_name' := 'cmp_rts_DFC_rbr_dsmtestErrorDFC'}
TYPE DFC_rbr_dsmtestErrorDFC : STRUCT
		DTC            : UDINT := 16#071200;
		DFCid          : UINT  := 881;
		debounceMethod : USINT := NO_DEBOUNCE;
	END_STRUCT
END_TYPE

(* ---- dfc_rbr_dsmupdatedeberror-DFC_rbr_dsmUpdateDebError.st ---- *)
(* --- Interface --- *)
{attribute 'external_name' := 'cmp_rts_DFC_rbr_dsmUpdateDebError'}
TYPE DFC_rbr_dsmUpdateDebError : STRUCT
		DTC            : UDINT := 16#070800;
		DFCid          : UINT  := 878;
		debounceMethod : USINT := NO_DEBOUNCE;
	END_STRUCT
END_TYPE

(* ---- dfc_rbr_dsmupdateerror-DFC_rbr_dsmUpdateError.st ---- *)
(* --- Interface --- *)
{attribute 'external_name' := 'cmp_rts_DFC_rbr_dsmUpdateError'}
TYPE DFC_rbr_dsmUpdateError : STRUCT
		DTC            : UDINT := 16#070900;
		DFCid          : UINT  := 879;
		debounceMethod : USINT := NO_DEBOUNCE;
	END_STRUCT
END_TYPE

(* ---- dfc_rbr_ina13or-DFC_rbr_inA13OR.st ---- *)
(* --- Interface --- *)
{attribute 'external_name' := 'cmp_rts_DFC_rbr_inA13OR'}
TYPE DFC_rbr_inA13OR : STRUCT
		DTC            : UDINT := 16#130100;
		DFCid          : UINT  := 209;
		debounceMethod : USINT := TIME_UP_DOWN;
	END_STRUCT
END_TYPE

(* ---- dfc_rbr_ina13scb-DFC_rbr_inA13SCB.st ---- *)
(* --- Interface --- *)
{attribute 'external_name' := 'cmp_rts_DFC_rbr_inA13SCB'}
TYPE DFC_rbr_inA13SCB : STRUCT
		DTC            : UDINT := 16#130200;
		DFCid          : UINT  := 210;
		debounceMethod : USINT := TIME_UP_DOWN;
	END_STRUCT
END_TYPE

(* ---- dfc_rbr_ina13scg-DFC_rbr_inA13SCG.st ---- *)
(* --- Interface --- *)
{attribute 'external_name' := 'cmp_rts_DFC_rbr_inA13SCG'}
TYPE DFC_rbr_inA13SCG : STRUCT
		DTC            : UDINT := 16#130300;
		DFCid          : UINT  := 211;
		debounceMethod : USINT := TIME_UP_DOWN;
	END_STRUCT
END_TYPE

(* ---- dfc_rbr_ina14or-DFC_rbr_inA14OR.st ---- *)
(* --- Interface --- *)
{attribute 'external_name' := 'cmp_rts_DFC_rbr_inA14OR'}
TYPE DFC_rbr_inA14OR : STRUCT
		DTC            : UDINT := 16#130400;
		DFCid          : UINT  := 212;
		debounceMethod : USINT := TIME_UP_DOWN;
	END_STRUCT
END_TYPE

(* ---- dfc_rbr_ina14scb-DFC_rbr_inA14SCB.st ---- *)
(* --- Interface --- *)
{attribute 'external_name' := 'cmp_rts_DFC_rbr_inA14SCB'}
TYPE DFC_rbr_inA14SCB : STRUCT
		DTC            : UDINT := 16#130500;
		DFCid          : UINT  := 213;
		debounceMethod : USINT := TIME_UP_DOWN;
	END_STRUCT
END_TYPE

(* ---- dfc_rbr_ina14scg-DFC_rbr_inA14SCG.st ---- *)
(* --- Interface --- *)
{attribute 'external_name' := 'cmp_rts_DFC_rbr_inA14SCG'}
TYPE DFC_rbr_inA14SCG : STRUCT
		DTC            : UDINT := 16#130600;
		DFCid          : UINT  := 214;
		debounceMethod : USINT := TIME_UP_DOWN;
	END_STRUCT
END_TYPE

(* ---- dfc_rbr_ina21or-DFC_rbr_inA21OR.st ---- *)
(* --- Interface --- *)
{attribute 'external_name' := 'cmp_rts_DFC_rbr_inA21OR'}
TYPE DFC_rbr_inA21OR : STRUCT
		DTC            : UDINT := 16#130700;
		DFCid          : UINT  := 215;
		debounceMethod : USINT := TIME_UP_DOWN;
	END_STRUCT
END_TYPE

(* ---- dfc_rbr_ina21scb-DFC_rbr_inA21SCB.st ---- *)
(* --- Interface --- *)
{attribute 'external_name' := 'cmp_rts_DFC_rbr_inA21SCB'}
TYPE DFC_rbr_inA21SCB : STRUCT
		DTC            : UDINT := 16#130800;
		DFCid          : UINT  := 216;
		debounceMethod : USINT := TIME_UP_DOWN;
	END_STRUCT
END_TYPE

(* ---- dfc_rbr_ina21scg-DFC_rbr_inA21SCG.st ---- *)
(* --- Interface --- *)
{attribute 'external_name' := 'cmp_rts_DFC_rbr_inA21SCG'}
TYPE DFC_rbr_inA21SCG : STRUCT
		DTC            : UDINT := 16#130900;
		DFCid          : UINT  := 217;
		debounceMethod : USINT := TIME_UP_DOWN;
	END_STRUCT
END_TYPE

(* ---- dfc_rbr_ina22or-DFC_rbr_inA22OR.st ---- *)
(* --- Interface --- *)
{attribute 'external_name' := 'cmp_rts_DFC_rbr_inA22OR'}
TYPE DFC_rbr_inA22OR : STRUCT
		DTC            : UDINT := 16#130A00;
		DFCid          : UINT  := 218;
		debounceMethod : USINT := TIME_UP_DOWN;
	END_STRUCT
END_TYPE

(* ---- dfc_rbr_ina22scb-DFC_rbr_inA22SCB.st ---- *)
(* --- Interface --- *)
{attribute 'external_name' := 'cmp_rts_DFC_rbr_inA22SCB'}
TYPE DFC_rbr_inA22SCB : STRUCT
		DTC            : UDINT := 16#130B00;
		DFCid          : UINT  := 219;
		debounceMethod : USINT := TIME_UP_DOWN;
	END_STRUCT
END_TYPE

(* ---- dfc_rbr_ina22scg-DFC_rbr_inA22SCG.st ---- *)
(* --- Interface --- *)
{attribute 'external_name' := 'cmp_rts_DFC_rbr_inA22SCG'}
TYPE DFC_rbr_inA22SCG : STRUCT
		DTC            : UDINT := 16#130C00;
		DFCid          : UINT  := 220;
		debounceMethod : USINT := TIME_UP_DOWN;
	END_STRUCT
END_TYPE

(* ---- dfc_rbr_ina23or-DFC_rbr_inA23OR.st ---- *)
(* --- Interface --- *)
{attribute 'external_name' := 'cmp_rts_DFC_rbr_inA23OR'}
TYPE DFC_rbr_inA23OR : STRUCT
		DTC            : UDINT := 16#130D00;
		DFCid          : UINT  := 221;
		debounceMethod : USINT := TIME_UP_DOWN;
	END_STRUCT
END_TYPE

(* ---- dfc_rbr_ina23scb-DFC_rbr_inA23SCB.st ---- *)
(* --- Interface --- *)
{attribute 'external_name' := 'cmp_rts_DFC_rbr_inA23SCB'}
TYPE DFC_rbr_inA23SCB : STRUCT
		DTC            : UDINT := 16#130E00;
		DFCid          : UINT  := 222;
		debounceMethod : USINT := TIME_UP_DOWN;
	END_STRUCT
END_TYPE

(* ---- dfc_rbr_ina23scg-DFC_rbr_inA23SCG.st ---- *)
(* --- Interface --- *)
{attribute 'external_name' := 'cmp_rts_DFC_rbr_inA23SCG'}
TYPE DFC_rbr_inA23SCG : STRUCT
		DTC            : UDINT := 16#130F00;
		DFCid          : UINT  := 223;
		debounceMethod : USINT := TIME_UP_DOWN;
	END_STRUCT
END_TYPE

(* ---- dfc_rbr_ina24or-DFC_rbr_inA24OR.st ---- *)
(* --- Interface --- *)
{attribute 'external_name' := 'cmp_rts_DFC_rbr_inA24OR'}
TYPE DFC_rbr_inA24OR : STRUCT
		DTC            : UDINT := 16#131000;
		DFCid          : UINT  := 224;
		debounceMethod : USINT := TIME_UP_DOWN;
	END_STRUCT
END_TYPE

(* ---- dfc_rbr_ina24scb-DFC_rbr_inA24SCB.st ---- *)
(* --- Interface --- *)
{attribute 'external_name' := 'cmp_rts_DFC_rbr_inA24SCB'}
TYPE DFC_rbr_inA24SCB : STRUCT
		DTC            : UDINT := 16#131100;
		DFCid          : UINT  := 225;
		debounceMethod : USINT := TIME_UP_DOWN;
	END_STRUCT
END_TYPE

(* ---- dfc_rbr_ina24scg-DFC_rbr_inA24SCG.st ---- *)
(* --- Interface --- *)
{attribute 'external_name' := 'cmp_rts_DFC_rbr_inA24SCG'}
TYPE DFC_rbr_inA24SCG : STRUCT
		DTC            : UDINT := 16#131200;
		DFCid          : UINT  := 226;
		debounceMethod : USINT := TIME_UP_DOWN;
	END_STRUCT
END_TYPE

(* ---- dfc_rbr_ina25or-DFC_rbr_inA25OR.st ---- *)
(* --- Interface --- *)
{attribute 'external_name' := 'cmp_rts_DFC_rbr_inA25OR'}
TYPE DFC_rbr_inA25OR : STRUCT
		DTC            : UDINT := 16#131300;
		DFCid          : UINT  := 227;
		debounceMethod : USINT := TIME_UP_DOWN;
	END_STRUCT
END_TYPE

(* ---- dfc_rbr_ina25scb-DFC_rbr_inA25SCB.st ---- *)
(* --- Interface --- *)
{attribute 'external_name' := 'cmp_rts_DFC_rbr_inA25SCB'}
TYPE DFC_rbr_inA25SCB : STRUCT
		DTC            : UDINT := 16#131400;
		DFCid          : UINT  := 228;
		debounceMethod : USINT := TIME_UP_DOWN;
	END_STRUCT
END_TYPE

(* ---- dfc_rbr_ina25scg-DFC_rbr_inA25SCG.st ---- *)
(* --- Interface --- *)
{attribute 'external_name' := 'cmp_rts_DFC_rbr_inA25SCG'}
TYPE DFC_rbr_inA25SCG : STRUCT
		DTC            : UDINT := 16#131500;
		DFCid          : UINT  := 229;
		debounceMethod : USINT := TIME_UP_DOWN;
	END_STRUCT
END_TYPE

(* ---- dfc_rbr_ina26or-DFC_rbr_inA26OR.st ---- *)
(* --- Interface --- *)
{attribute 'external_name' := 'cmp_rts_DFC_rbr_inA26OR'}
TYPE DFC_rbr_inA26OR : STRUCT
		DTC            : UDINT := 16#131600;
		DFCid          : UINT  := 230;
		debounceMethod : USINT := TIME_UP_DOWN;
	END_STRUCT
END_TYPE

(* ---- dfc_rbr_ina26scb-DFC_rbr_inA26SCB.st ---- *)
(* --- Interface --- *)
{attribute 'external_name' := 'cmp_rts_DFC_rbr_inA26SCB'}
TYPE DFC_rbr_inA26SCB : STRUCT
		DTC            : UDINT := 16#131700;
		DFCid          : UINT  := 231;
		debounceMethod : USINT := TIME_UP_DOWN;
	END_STRUCT
END_TYPE

(* ---- dfc_rbr_ina26scg-DFC_rbr_inA26SCG.st ---- *)
(* --- Interface --- *)
{attribute 'external_name' := 'cmp_rts_DFC_rbr_inA26SCG'}
TYPE DFC_rbr_inA26SCG : STRUCT
		DTC            : UDINT := 16#131800;
		DFCid          : UINT  := 232;
		debounceMethod : USINT := TIME_UP_DOWN;
	END_STRUCT
END_TYPE

(* ---- dfc_rbr_ina27or-DFC_rbr_inA27OR.st ---- *)
(* --- Interface --- *)
{attribute 'external_name' := 'cmp_rts_DFC_rbr_inA27OR'}
TYPE DFC_rbr_inA27OR : STRUCT
		DTC            : UDINT := 16#131900;
		DFCid          : UINT  := 233;
		debounceMethod : USINT := TIME_UP_DOWN;
	END_STRUCT
END_TYPE

(* ---- dfc_rbr_ina27scb-DFC_rbr_inA27SCB.st ---- *)
(* --- Interface --- *)
{attribute 'external_name' := 'cmp_rts_DFC_rbr_inA27SCB'}
TYPE DFC_rbr_inA27SCB : STRUCT
		DTC            : UDINT := 16#131A00;
		DFCid          : UINT  := 234;
		debounceMethod : USINT := TIME_UP_DOWN;
	END_STRUCT
END_TYPE

(* ---- dfc_rbr_ina27scg-DFC_rbr_inA27SCG.st ---- *)
(* --- Interface --- *)
{attribute 'external_name' := 'cmp_rts_DFC_rbr_inA27SCG'}
TYPE DFC_rbr_inA27SCG : STRUCT
		DTC            : UDINT := 16#131B00;
		DFCid          : UINT  := 235;
		debounceMethod : USINT := TIME_UP_DOWN;
	END_STRUCT
END_TYPE

(* ---- dfc_rbr_ina28or-DFC_rbr_inA28OR.st ---- *)
(* --- Interface --- *)
{attribute 'external_name' := 'cmp_rts_DFC_rbr_inA28OR'}
TYPE DFC_rbr_inA28OR : STRUCT
		DTC            : UDINT := 16#131C00;
		DFCid          : UINT  := 236;
		debounceMethod : USINT := TIME_UP_DOWN;
	END_STRUCT
END_TYPE

(* ---- dfc_rbr_ina28scb-DFC_rbr_inA28SCB.st ---- *)
(* --- Interface --- *)
{attribute 'external_name' := 'cmp_rts_DFC_rbr_inA28SCB'}
TYPE DFC_rbr_inA28SCB : STRUCT
		DTC            : UDINT := 16#131D00;
		DFCid          : UINT  := 237;
		debounceMethod : USINT := TIME_UP_DOWN;
	END_STRUCT
END_TYPE

(* ---- dfc_rbr_ina28scg-DFC_rbr_inA28SCG.st ---- *)
(* --- Interface --- *)
{attribute 'external_name' := 'cmp_rts_DFC_rbr_inA28SCG'}
TYPE DFC_rbr_inA28SCG : STRUCT
		DTC            : UDINT := 16#131E00;
		DFCid          : UINT  := 238;
		debounceMethod : USINT := TIME_UP_DOWN;
	END_STRUCT
END_TYPE

(* ---- dfc_rbr_ina29or-DFC_rbr_inA29OR.st ---- *)
(* --- Interface --- *)
{attribute 'external_name' := 'cmp_rts_DFC_rbr_inA29OR'}
TYPE DFC_rbr_inA29OR : STRUCT
		DTC            : UDINT := 16#131F00;
		DFCid          : UINT  := 239;
		debounceMethod : USINT := TIME_UP_DOWN;
	END_STRUCT
END_TYPE

(* ---- dfc_rbr_ina29scb-DFC_rbr_inA29SCB.st ---- *)
(* --- Interface --- *)
{attribute 'external_name' := 'cmp_rts_DFC_rbr_inA29SCB'}
TYPE DFC_rbr_inA29SCB : STRUCT
		DTC            : UDINT := 16#132000;
		DFCid          : UINT  := 240;
		debounceMethod : USINT := TIME_UP_DOWN;
	END_STRUCT
END_TYPE

(* ---- dfc_rbr_ina29scg-DFC_rbr_inA29SCG.st ---- *)
(* --- Interface --- *)
{attribute 'external_name' := 'cmp_rts_DFC_rbr_inA29SCG'}
TYPE DFC_rbr_inA29SCG : STRUCT
		DTC            : UDINT := 16#132100;
		DFCid          : UINT  := 241;
		debounceMethod : USINT := TIME_UP_DOWN;
	END_STRUCT
END_TYPE

(* ---- dfc_rbr_ina36aicscb-DFC_rbr_inA36AicSCB.st ---- *)
(* --- Interface --- *)
{attribute 'external_name' := 'cmp_rts_DFC_rbr_inA36AicSCB'}
TYPE DFC_rbr_inA36AicSCB : STRUCT
		DTC            : UDINT := 16#132200;
		DFCid          : UINT  := 242;
		debounceMethod : USINT := TIME_UP_DOWN;
	END_STRUCT
END_TYPE

(* ---- dfc_rbr_ina36aicscg-DFC_rbr_inA36AicSCG.st ---- *)
(* --- Interface --- *)
{attribute 'external_name' := 'cmp_rts_DFC_rbr_inA36AicSCG'}
TYPE DFC_rbr_inA36AicSCG : STRUCT
		DTC            : UDINT := 16#132300;
		DFCid          : UINT  := 243;
		debounceMethod : USINT := TIME_UP_DOWN;
	END_STRUCT
END_TYPE

(* ---- dfc_rbr_ina36or-DFC_rbr_inA36OR.st ---- *)
(* --- Interface --- *)
{attribute 'external_name' := 'cmp_rts_DFC_rbr_inA36OR'}
TYPE DFC_rbr_inA36OR : STRUCT
		DTC            : UDINT := 16#132400;
		DFCid          : UINT  := 244;
		debounceMethod : USINT := TIME_UP_DOWN;
	END_STRUCT
END_TYPE

(* ---- dfc_rbr_ina36scb-DFC_rbr_inA36SCB.st ---- *)
(* --- Interface --- *)
{attribute 'external_name' := 'cmp_rts_DFC_rbr_inA36SCB'}
TYPE DFC_rbr_inA36SCB : STRUCT
		DTC            : UDINT := 16#132500;
		DFCid          : UINT  := 245;
		debounceMethod : USINT := TIME_UP_DOWN;
	END_STRUCT
END_TYPE

(* ---- dfc_rbr_ina36scg-DFC_rbr_inA36SCG.st ---- *)
(* --- Interface --- *)
{attribute 'external_name' := 'cmp_rts_DFC_rbr_inA36SCG'}
TYPE DFC_rbr_inA36SCG : STRUCT
		DTC            : UDINT := 16#132600;
		DFCid          : UINT  := 246;
		debounceMethod : USINT := TIME_UP_DOWN;
	END_STRUCT
END_TYPE

(* ---- dfc_rbr_ina36shuntscb-DFC_rbr_inA36ShuntSCB.st ---- *)
(* --- Interface --- *)
{attribute 'external_name' := 'cmp_rts_DFC_rbr_inA36ShuntSCB'}
TYPE DFC_rbr_inA36ShuntSCB : STRUCT
		DTC            : UDINT := 16#132700;
		DFCid          : UINT  := 247;
		debounceMethod : USINT := TIME_UP_DOWN;
	END_STRUCT
END_TYPE

(* ---- dfc_rbr_ina37aicscb-DFC_rbr_inA37AicSCB.st ---- *)
(* --- Interface --- *)
{attribute 'external_name' := 'cmp_rts_DFC_rbr_inA37AicSCB'}
TYPE DFC_rbr_inA37AicSCB : STRUCT
		DTC            : UDINT := 16#132800;
		DFCid          : UINT  := 248;
		debounceMethod : USINT := TIME_UP_DOWN;
	END_STRUCT
END_TYPE

(* ---- dfc_rbr_ina37aicscg-DFC_rbr_inA37AicSCG.st ---- *)
(* --- Interface --- *)
{attribute 'external_name' := 'cmp_rts_DFC_rbr_inA37AicSCG'}
TYPE DFC_rbr_inA37AicSCG : STRUCT
		DTC            : UDINT := 16#132900;
		DFCid          : UINT  := 249;
		debounceMethod : USINT := TIME_UP_DOWN;
	END_STRUCT
END_TYPE

(* ---- dfc_rbr_ina37or-DFC_rbr_inA37OR.st ---- *)
(* --- Interface --- *)
{attribute 'external_name' := 'cmp_rts_DFC_rbr_inA37OR'}
TYPE DFC_rbr_inA37OR : STRUCT
		DTC            : UDINT := 16#132A00;
		DFCid          : UINT  := 250;
		debounceMethod : USINT := TIME_UP_DOWN;
	END_STRUCT
END_TYPE

(* ---- dfc_rbr_ina37scb-DFC_rbr_inA37SCB.st ---- *)
(* --- Interface --- *)
{attribute 'external_name' := 'cmp_rts_DFC_rbr_inA37SCB'}
TYPE DFC_rbr_inA37SCB : STRUCT
		DTC            : UDINT := 16#132B00;
		DFCid          : UINT  := 251;
		debounceMethod : USINT := TIME_UP_DOWN;
	END_STRUCT
END_TYPE

(* ---- dfc_rbr_ina37scg-DFC_rbr_inA37SCG.st ---- *)
(* --- Interface --- *)
{attribute 'external_name' := 'cmp_rts_DFC_rbr_inA37SCG'}
TYPE DFC_rbr_inA37SCG : STRUCT
		DTC            : UDINT := 16#132C00;
		DFCid          : UINT  := 252;
		debounceMethod : USINT := TIME_UP_DOWN;
	END_STRUCT
END_TYPE

(* ---- dfc_rbr_ina37shuntscb-DFC_rbr_inA37ShuntSCB.st ---- *)
(* --- Interface --- *)
{attribute 'external_name' := 'cmp_rts_DFC_rbr_inA37ShuntSCB'}
TYPE DFC_rbr_inA37ShuntSCB : STRUCT
		DTC            : UDINT := 16#132D00;
		DFCid          : UINT  := 253;
		debounceMethod : USINT := TIME_UP_DOWN;
	END_STRUCT
END_TYPE

(* ---- dfc_rbr_ina38aicscb-DFC_rbr_inA38AicSCB.st ---- *)
(* --- Interface --- *)
{attribute 'external_name' := 'cmp_rts_DFC_rbr_inA38AicSCB'}
TYPE DFC_rbr_inA38AicSCB : STRUCT
		DTC            : UDINT := 16#132E00;
		DFCid          : UINT  := 254;
		debounceMethod : USINT := TIME_UP_DOWN;
	END_STRUCT
END_TYPE

(* ---- dfc_rbr_ina38aicscg-DFC_rbr_inA38AicSCG.st ---- *)
(* --- Interface --- *)
{attribute 'external_name' := 'cmp_rts_DFC_rbr_inA38AicSCG'}
TYPE DFC_rbr_inA38AicSCG : STRUCT
		DTC            : UDINT := 16#132F00;
		DFCid          : UINT  := 255;
		debounceMethod : USINT := TIME_UP_DOWN;
	END_STRUCT
END_TYPE

(* ---- dfc_rbr_ina38or-DFC_rbr_inA38OR.st ---- *)
(* --- Interface --- *)
{attribute 'external_name' := 'cmp_rts_DFC_rbr_inA38OR'}
TYPE DFC_rbr_inA38OR : STRUCT
		DTC            : UDINT := 16#133000;
		DFCid          : UINT  := 256;
		debounceMethod : USINT := TIME_UP_DOWN;
	END_STRUCT
END_TYPE
